REGION Network 16: Step7: Request Take Photos and Calculate Again When ROS Error | PLC Status Word:111 0r 112
   RUNG wire#powerrail
      Contact( #High )
      Contact( "DB2500 Visual Chiseling".VisualChiselingMode )
      Contact( "DB2500 Visual Chiseling".VisualCameraStart )
      wire#w1
      { S7_Templates := "SrcType := Int" } EQ_Contact(in1 := "DB2500 Visual Chiseling".RosErrorNum, in2 := 1)
      P_Trig( "DB2500 Visual Chiseling".Pulse[9] )
      Move(in := 111, out1 => "DB2100 Modbus Value"."PLC Para"."Status Word")
   END_RUNG
   RUNG wire#w1
      { S7_Templates := "SrcType := Int" } EQ_Contact(in1 := "DB2500 Visual Chiseling".RosErrorNum, in2 := 2)
      P_Trig( "DB2500 Visual Chiseling".Pulse[10] )
      Move(in := 112, out1 => "DB2100 Modbus Value"."PLC Para"."Status Word")
   END_RUNG
   // the same network as SCL:
   #_w1 := #High AND "DB2500 Visual Chiseling".VisualChiselingMode AND "DB2500 Visual Chiseling".VisualCameraStart;
   #_w2 := #_w1 AND ("DB2500 Visual Chiseling".RosErrorNum = 1);
   #_w3 := #_w2 AND NOT "DB2500 Visual Chiseling".Pulse[9];   // rising edge
   "DB2500 Visual Chiseling".Pulse[9] := #_w2;
   IF #_w3 THEN "DB2100 Modbus Value"."PLC Para"."Status Word" := 111; END_IF;
   #_w4 := #_w1 AND ("DB2500 Visual Chiseling".RosErrorNum = 2);
   #_w5 := #_w4 AND NOT "DB2500 Visual Chiseling".Pulse[10];   // rising edge
   "DB2500 Visual Chiseling".Pulse[10] := #_w4;
   IF #_w5 THEN "DB2100 Modbus Value"."PLC Para"."Status Word" := 112; END_IF;
END_REGION

REGION Network 17: Step7: Stop Communication and SShutDown ROS If Erro Num Bigger Than 3 | PLC Status Word:105
   // Status 105: Send Shut Down Signal to ROS
   RUNG wire#powerrail
      Contact( #High )
      Contact( "DB2500 Visual Chiseling".VisualChiselingMode )
      Contact( "DB2500 Visual Chiseling".VisualCameraStart )
      { S7_Templates := "SrcType := Int" } GE_Contact(in1 := "DB2500 Visual Chiseling".RosErrorNum, in2 := 3)
      P_Trig( "DB2500 Visual Chiseling".Pulse[11] )
      wire#w1
      Move(in := 105, out1 => "DB2100 Modbus Value"."PLC Para"."Status Word")
   END_RUNG
   RUNG wire#w1
      S_Coil( "DB2500 Visual Chiseling".ROSCalculationFault )
      R_Coil( "DB2500 Visual Chiseling".VisualCameraStart )
   END_RUNG
   // the same network as SCL:
   #_w1 := #High AND "DB2500 Visual Chiseling".VisualChiselingMode AND "DB2500 Visual Chiseling".VisualCameraStart AND ("DB2500 Visual Chiseling".RosErrorNum >= 3);
   #_w2 := #_w1 AND NOT "DB2500 Visual Chiseling".Pulse[11];   // rising edge
   "DB2500 Visual Chiseling".Pulse[11] := #_w1;
   IF #_w2 THEN
       "DB2100 Modbus Value"."PLC Para"."Status Word" := 105;
       "DB2500 Visual Chiseling".ROSCalculationFault := TRUE;
       "DB2500 Visual Chiseling".VisualCameraStart := FALSE;
   END_IF;
END_REGION

REGION Network 18: Step8: Auto Close Camera Protective Cover | PLC Status Word:130
   "Timer30_ChiselStepEnd".TON(IN := #High AND "DB2500 Visual Chiseling".VisualChiselingMode AND "DB2500 Visual Chiseling".VisualCameraStart AND (("DB2100 Modbus Value"."PLC Para"."Status Word" = 120) OR "DB2500 Visual Chiseling".ROSCalculationFault),
                           PT := T#0.2s);
   IF "Timer30_ChiselStepEnd".Q THEN "DB2100 Modbus Value"."PLC Para"."Status Word" := 130; END_IF;
END_REGION

REGION Network 19: Step9: Visual Chiseling Camera Function Completed
   // Robot: IN[80]   PLC :DB720.DBX2.0  VisualChiseling  Camera Function  Completion Signal
   RUNG wire#powerrail
      Contact( #High )
      Contact( "DB2500 Visual Chiseling".VisualChiselingMode )
      Contact( "DB2500 Visual Chiseling".VisualCameraStart )
      { S7_Templates := "SrcType := Word" } EQ_Contact(in1 := "DB2100 Modbus Value"."PLC Para"."Status Word", in2 := 130)
      P_Trig( "DB2500 Visual Chiseling".Pulse[12] )
      wire#w1
      Move(in := 0, out1 => "DB2500 Visual Chiseling".RosErrorNum)
   END_RUNG
   RUNG wire#w1
      R_Coil( "DB2500 Visual Chiseling".VisualCameraStart )
      S_Coil( "DB2500 Visual Chiseling".VisualCameraEnd )
      R_Coil( "QCamCoverExt" )
      S_Coil( "QCamCoverRet" )
   END_RUNG
   // the same network as SCL:
   #_w1 := #High AND "DB2500 Visual Chiseling".VisualChiselingMode AND "DB2500 Visual Chiseling".VisualCameraStart AND ("DB2100 Modbus Value"."PLC Para"."Status Word" = 130);
   #_w2 := #_w1 AND NOT "DB2500 Visual Chiseling".Pulse[12];   // rising edge
   "DB2500 Visual Chiseling".Pulse[12] := #_w1;
   IF #_w2 THEN
       "DB2500 Visual Chiseling".RosErrorNum := 0;
       "DB2500 Visual Chiseling".VisualCameraStart := FALSE;
       "DB2500 Visual Chiseling".VisualCameraEnd := TRUE;
       "QCamCoverExt" := FALSE;
       "QCamCoverRet" := TRUE;
   END_IF;
END_REGION

REGION Network 20: Step9.1 : Send Visual Chiseling Function Completion Signal to Robot.
   // Robot: IN[80]   PLC :DB720.DBX2.0  VisualChiseling  Camera Function  Completion Signal
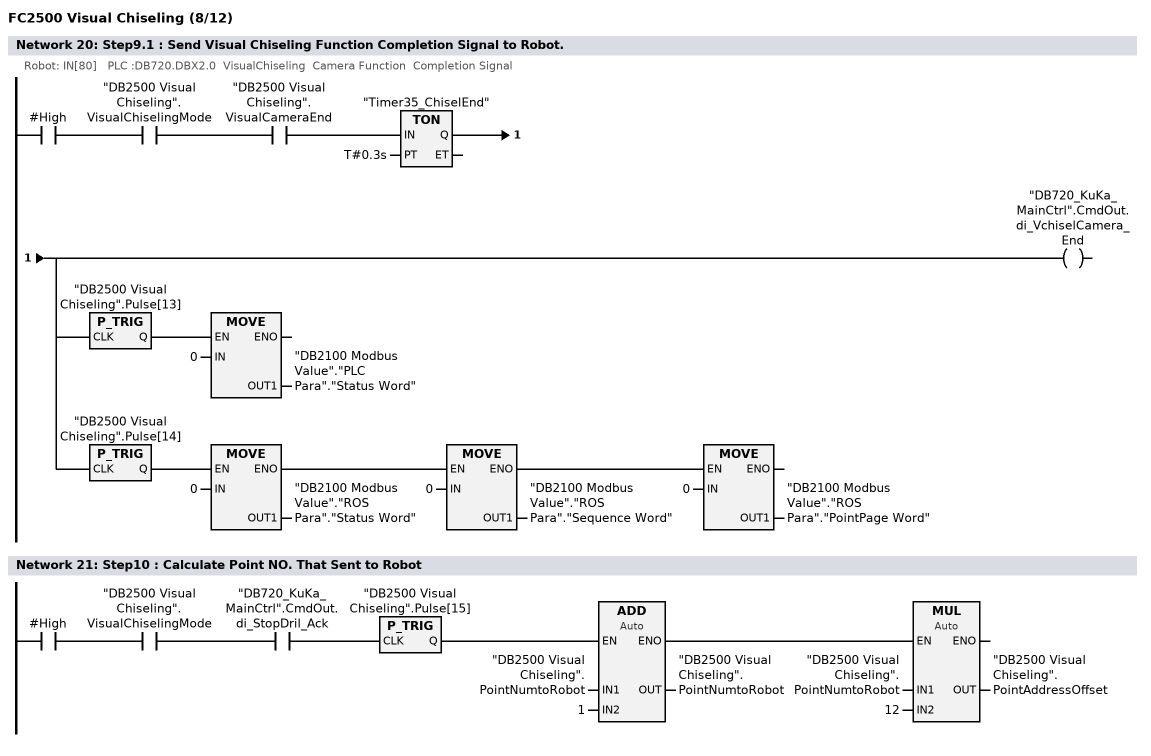
   "Timer35_ChiselEnd".TON(IN := #High AND "DB2500 Visual Chiseling".VisualChiselingMode AND "DB2500 Visual Chiseling".VisualCameraEnd,
                           PT := T#0.3s);
   "DB720_KuKa_MainCtrl".CmdOut.di_VchiselCamera_End := "Timer35_ChiselEnd".Q;
   #_w1 := "Timer35_ChiselEnd".Q AND NOT "DB2500 Visual Chiseling".Pulse[13];   // rising edge
   "DB2500 Visual Chiseling".Pulse[13] := "Timer35_ChiselEnd".Q;
   IF #_w1 THEN "DB2100 Modbus Value"."PLC Para"."Status Word" := 0; END_IF;
   #_w2 := "Timer35_ChiselEnd".Q AND NOT "DB2500 Visual Chiseling".Pulse[14];   // rising edge
   "DB2500 Visual Chiseling".Pulse[14] := "Timer35_ChiselEnd".Q;
   IF #_w2 THEN
       "DB2100 Modbus Value"."ROS Para"."Status Word" := 0;
       "DB2100 Modbus Value"."ROS Para"."Sequence Word" := 0;
       "DB2100 Modbus Value"."ROS Para"."PointPage Word" := 0;
   END_IF;
END_REGION

REGION Network 21: Step10 : Calculate Point NO. That Sent to Robot
   RUNG wire#powerrail
      Contact( #High )
      Contact( "DB2500 Visual Chiseling".VisualChiselingMode )
      Contact( "DB720_KuKa_MainCtrl".CmdOut.di_StopDril_Ack )
      P_Trig( "DB2500 Visual Chiseling".Pulse[15] )
      Add(in1 := "DB2500 Visual Chiseling".PointNumtoRobot, in2 := 1, out => "DB2500 Visual Chiseling".PointNumtoRobot)
      Mul(in1 := "DB2500 Visual Chiseling".PointNumtoRobot, in2 := 12, out => "DB2500 Visual Chiseling".PointAddressOffset)
   END_RUNG
   // the same network as SCL:
   #_w1 := #High AND "DB2500 Visual Chiseling".VisualChiselingMode AND "DB720_KuKa_MainCtrl".CmdOut.di_StopDril_Ack;
   #_w2 := #_w1 AND NOT "DB2500 Visual Chiseling".Pulse[15];   // rising edge
   "DB2500 Visual Chiseling".Pulse[15] := #_w1;
   IF #_w2 THEN
       "DB2500 Visual Chiseling".PointNumtoRobot := "DB2500 Visual Chiseling".PointNumtoRobot + 1;
       "DB2500 Visual Chiseling".PointAddressOffset := "DB2500 Visual Chiseling".PointNumtoRobot * 12;
   END_IF;
END_REGION

REGION Network 22 (SCL): Step11: Move Current Chiseling Point to Offset Value. (SCL)
   // byteOffset_dest Should Be Changed wehn
   IF "DB2500 Visual Chiseling".VisualCameraEnd = TRUE THEN
       POKE_BLK(area_src := 16#84,
                dbNumber_src := 2300,
                byteOffset_src := "DB2500 Visual Chiseling".PointAddressOffset,
                area_dest := 16#84,
                dbNumber_dest := 2500,
                byteOffset_dest := 38,
                count := 12);
   END_IF;
END_REGION

REGION Network 23: Step12: Offset Value Format From Word To Real
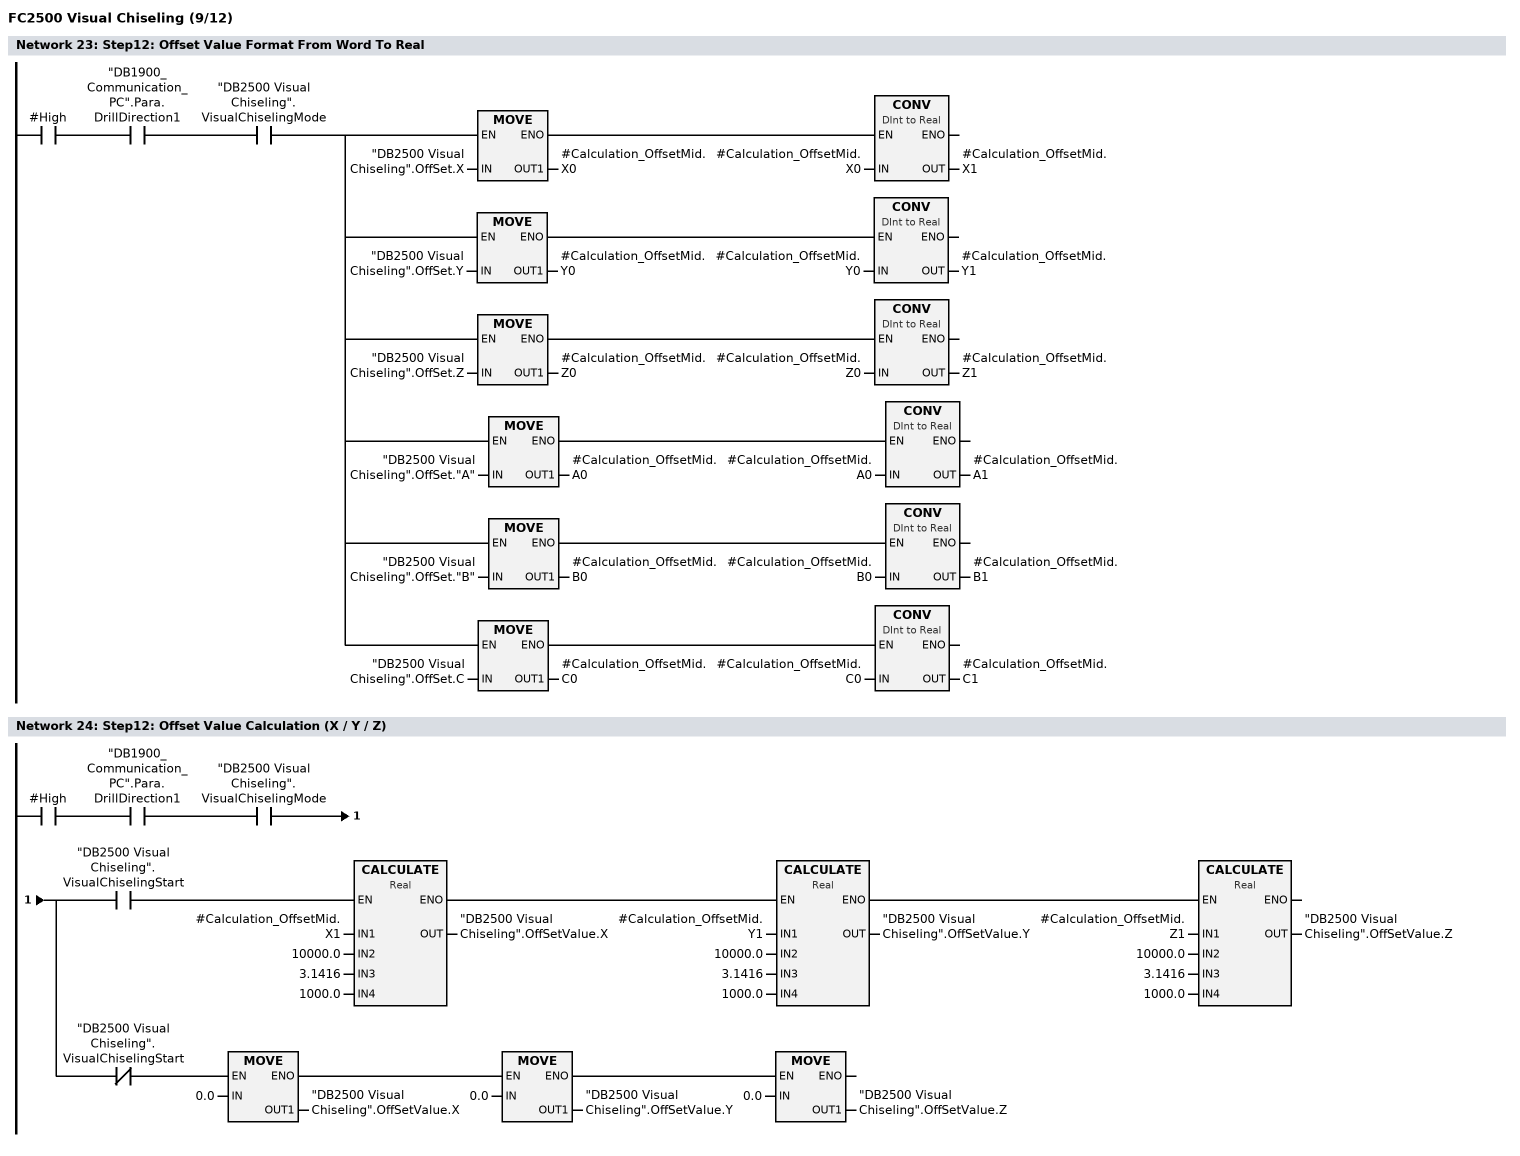
   RUNG wire#powerrail
      Contact( #High )
      Contact( "DB1900_Communication_PC".Para.DrillDirection1 )
      Contact( "DB2500 Visual Chiseling".VisualChiselingMode )
      wire#w1
      Move(in := "DB2500 Visual Chiseling".OffSet.X, out1 => #Calculation_OffsetMid.X0)
      { S7_Templates := "[SrcType := DInt, DestType := Real]" } Convert(in := #Calculation_OffsetMid.X0, out => #Calculation_OffsetMid.X1)
   END_RUNG
   RUNG wire#w1
      Move(in := "DB2500 Visual Chiseling".OffSet.Y, out1 => #Calculation_OffsetMid.Y0)
      { S7_Templates := "[SrcType := DInt, DestType := Real]" } Convert(in := #Calculation_OffsetMid.Y0, out => #Calculation_OffsetMid.Y1)
   END_RUNG
   RUNG wire#w1
      Move(in := "DB2500 Visual Chiseling".OffSet.Z, out1 => #Calculation_OffsetMid.Z0)
      { S7_Templates := "[SrcType := DInt, DestType := Real]" } Convert(in := #Calculation_OffsetMid.Z0, out => #Calculation_OffsetMid.Z1)
   END_RUNG
   RUNG wire#w1
      Move(in := "DB2500 Visual Chiseling".OffSet."A", out1 => #Calculation_OffsetMid.A0)
      { S7_Templates := "[SrcType := DInt, DestType := Real]" } Convert(in := #Calculation_OffsetMid.A0, out => #Calculation_OffsetMid.A1)
   END_RUNG
   RUNG wire#w1
      Move(in := "DB2500 Visual Chiseling".OffSet."B", out1 => #Calculation_OffsetMid.B0)
      { S7_Templates := "[SrcType := DInt, DestType := Real]" } Convert(in := #Calculation_OffsetMid.B0, out => #Calculation_OffsetMid.B1)
   END_RUNG
   RUNG wire#w1
      Move(in := "DB2500 Visual Chiseling".OffSet.C, out1 => #Calculation_OffsetMid.C0)
      { S7_Templates := "[SrcType := DInt, DestType := Real]" } Convert(in := #Calculation_OffsetMid.C0, out => #Calculation_OffsetMid.C1)
   END_RUNG
   // the same network as SCL:
   IF #High AND "DB1900_Communication_PC".Para.DrillDirection1 AND "DB2500 Visual Chiseling".VisualChiselingMode THEN
       #Calculation_OffsetMid.X0 := "DB2500 Visual Chiseling".OffSet.X;
       #Calculation_OffsetMid.X1 := DINT_TO_REAL(#Calculation_OffsetMid.X0);
       #Calculation_OffsetMid.Y0 := "DB2500 Visual Chiseling".OffSet.Y;
       #Calculation_OffsetMid.Y1 := DINT_TO_REAL(#Calculation_OffsetMid.Y0);
       #Calculation_OffsetMid.Z0 := "DB2500 Visual Chiseling".OffSet.Z;
       #Calculation_OffsetMid.Z1 := DINT_TO_REAL(#Calculation_OffsetMid.Z0);
       #Calculation_OffsetMid.A0 := "DB2500 Visual Chiseling".OffSet."A";
       #Calculation_OffsetMid.A1 := DINT_TO_REAL(#Calculation_OffsetMid.A0);
       #Calculation_OffsetMid.B0 := "DB2500 Visual Chiseling".OffSet."B";
       #Calculation_OffsetMid.B1 := DINT_TO_REAL(#Calculation_OffsetMid.B0);
       #Calculation_OffsetMid.C0 := "DB2500 Visual Chiseling".OffSet.C;
       #Calculation_OffsetMid.C1 := DINT_TO_REAL(#Calculation_OffsetMid.C0);
   END_IF;
END_REGION

REGION Network 24: Step12: Offset Value Calculation (X / Y / Z)
   RUNG wire#powerrail
      Contact( #High )
      Contact( "DB1900_Communication_PC".Para.DrillDirection1 )
      Contact( "DB2500 Visual Chiseling".VisualChiselingMode )
      wire#w1
      Contact( "DB2500 Visual Chiseling".VisualChiselingStart )
      { S7_Templates := "SrcType := Real"; S7_Expression := "( IN1 / IN2 - IN3 ) * IN4" } Calculate(in1 := #Calculation_OffsetMid.X1, in2 := 10000.0, in3 := 3.1416, in4 := 1000.0, out => "DB2500 Visual Chiseling".OffSetValue.X)
      { S7_Templates := "SrcType := Real"; S7_Expression := "( IN1 / IN2 - IN3 ) * IN4" } Calculate(in1 := #Calculation_OffsetMid.Y1, in2 := 10000.0, in3 := 3.1416, in4 := 1000.0, out => "DB2500 Visual Chiseling".OffSetValue.Y)
      { S7_Templates := "SrcType := Real"; S7_Expression := "( IN1 / IN2 - IN3 ) * IN4" } Calculate(in1 := #Calculation_OffsetMid.Z1, in2 := 10000.0, in3 := 3.1416, in4 := 1000.0, out => "DB2500 Visual Chiseling".OffSetValue.Z)
   END_RUNG
   RUNG wire#w1
      I_Contact( "DB2500 Visual Chiseling".VisualChiselingStart )
      Move(in := 0.0, out1 => "DB2500 Visual Chiseling".OffSetValue.X)
      Move(in := 0.0, out1 => "DB2500 Visual Chiseling".OffSetValue.Y)
      Move(in := 0.0, out1 => "DB2500 Visual Chiseling".OffSetValue.Z)
   END_RUNG
   // the same network as SCL:
   #_w1 := #High AND "DB1900_Communication_PC".Para.DrillDirection1 AND "DB2500 Visual Chiseling".VisualChiselingMode;
   IF #_w1 AND "DB2500 Visual Chiseling".VisualChiselingStart THEN
       "DB2500 Visual Chiseling".OffSetValue.X := ( #Calculation_OffsetMid.X1 / 10000.0 - 3.1416 ) * 1000.0;
       "DB2500 Visual Chiseling".OffSetValue.Y := ( #Calculation_OffsetMid.Y1 / 10000.0 - 3.1416 ) * 1000.0;
       "DB2500 Visual Chiseling".OffSetValue.Z := ( #Calculation_OffsetMid.Z1 / 10000.0 - 3.1416 ) * 1000.0;
   END_IF;
   IF #_w1 AND NOT "DB2500 Visual Chiseling".VisualChiselingStart THEN
       "DB2500 Visual Chiseling".OffSetValue.X := 0.0;
       "DB2500 Visual Chiseling".OffSetValue.Y := 0.0;
       "DB2500 Visual Chiseling".OffSetValue.Z := 0.0;
   END_IF;
END_REGION

REGION Network 25: Step13: Offset Value Calculation (A / B / C)
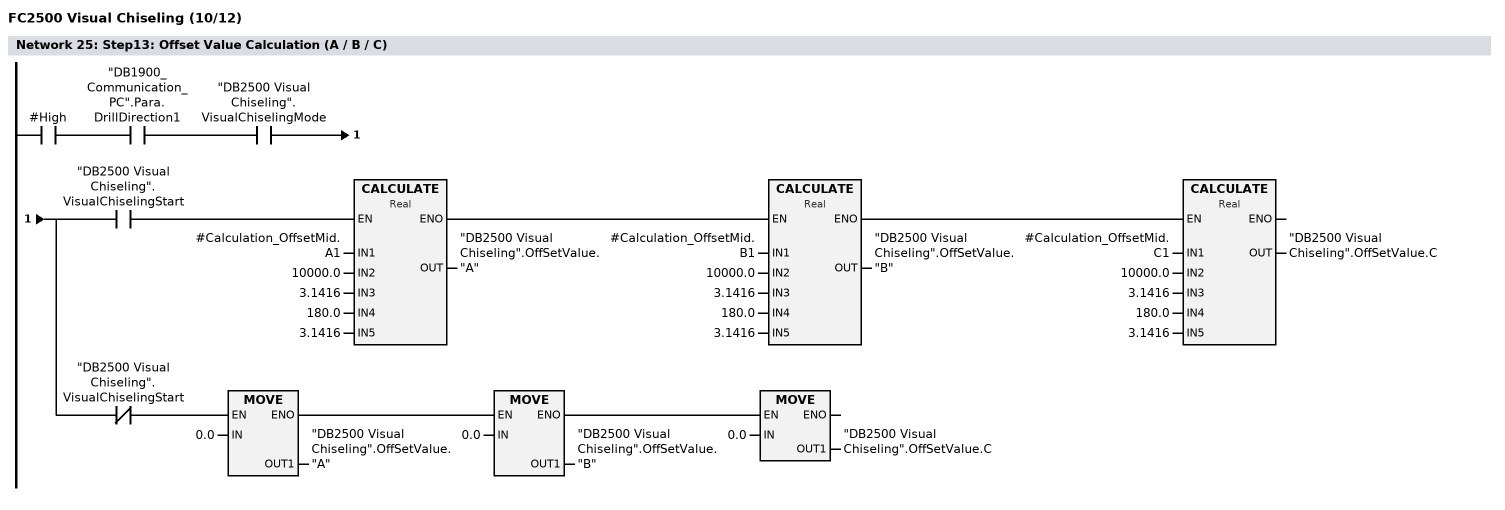
   RUNG wire#powerrail
      Contact( #High )
      Contact( "DB1900_Communication_PC".Para.DrillDirection1 )
      Contact( "DB2500 Visual Chiseling".VisualChiselingMode )
      wire#w1
      Contact( "DB2500 Visual Chiseling".VisualChiselingStart )
      { S7_Templates := "SrcType := Real"; S7_Expression := "( ( IN1 / IN2 - IN3 ) * IN4 ) / IN5" } Calculate(in1 := #Calculation_OffsetMid.A1, in2 := 10000.0, in3 := 3.1416, in4 := 180.0, in5 := 3.1416, out => "DB2500 Visual Chiseling".OffSetValue."A")
      { S7_Templates := "SrcType := Real"; S7_Expression := "( ( IN1 / IN2 - IN3 ) * IN4 ) / IN5" } Calculate(in1 := #Calculation_OffsetMid.B1, in2 := 10000.0, in3 := 3.1416, in4 := 180.0, in5 := 3.1416, out => "DB2500 Visual Chiseling".OffSetValue."B")
      { S7_Templates := "SrcType := Real"; S7_Expression := "( ( IN1 / IN2 - IN3 ) * IN4 ) / IN5" } Calculate(in1 := #Calculation_OffsetMid.C1, in2 := 10000.0, in3 := 3.1416, in4 := 180.0, in5 := 3.1416, out => "DB2500 Visual Chiseling".OffSetValue.C)
   END_RUNG
   RUNG wire#w1
      I_Contact( "DB2500 Visual Chiseling".VisualChiselingStart )
      Move(in := 0.0, out1 => "DB2500 Visual Chiseling".OffSetValue."A")
      Move(in := 0.0, out1 => "DB2500 Visual Chiseling".OffSetValue."B")
      Move(in := 0.0, out1 => "DB2500 Visual Chiseling".OffSetValue.C)
   END_RUNG
   // the same network as SCL:
   #_w1 := #High AND "DB1900_Communication_PC".Para.DrillDirection1 AND "DB2500 Visual Chiseling".VisualChiselingMode;
   IF #_w1 AND "DB2500 Visual Chiseling".VisualChiselingStart THEN
       "DB2500 Visual Chiseling".OffSetValue."A" := ( ( #Calculation_OffsetMid.A1 / 10000.0 - 3.1416 ) * 180.0 ) / 3.1416;
       "DB2500 Visual Chiseling".OffSetValue."B" := ( ( #Calculation_OffsetMid.B1 / 10000.0 - 3.1416 ) * 180.0 ) / 3.1416;
       "DB2500 Visual Chiseling".OffSetValue.C := ( ( #Calculation_OffsetMid.C1 / 10000.0 - 3.1416 ) * 180.0 ) / 3.1416;
   END_IF;
   IF #_w1 AND NOT "DB2500 Visual Chiseling".VisualChiselingStart THEN
       "DB2500 Visual Chiseling".OffSetValue."A" := 0.0;
       "DB2500 Visual Chiseling".OffSetValue."B" := 0.0;
       "DB2500 Visual Chiseling".OffSetValue.C := 0.0;
   END_IF;
END_REGION

REGION Network 26: Step14: Transfer Offset Value to Robot
   // Added by WXY 20220618.  DBD720.DBD36: gi_OffSetA;  DBD720.DBD40: gi_OffSetB;   DBD720.DBD44: gi_OffSetC
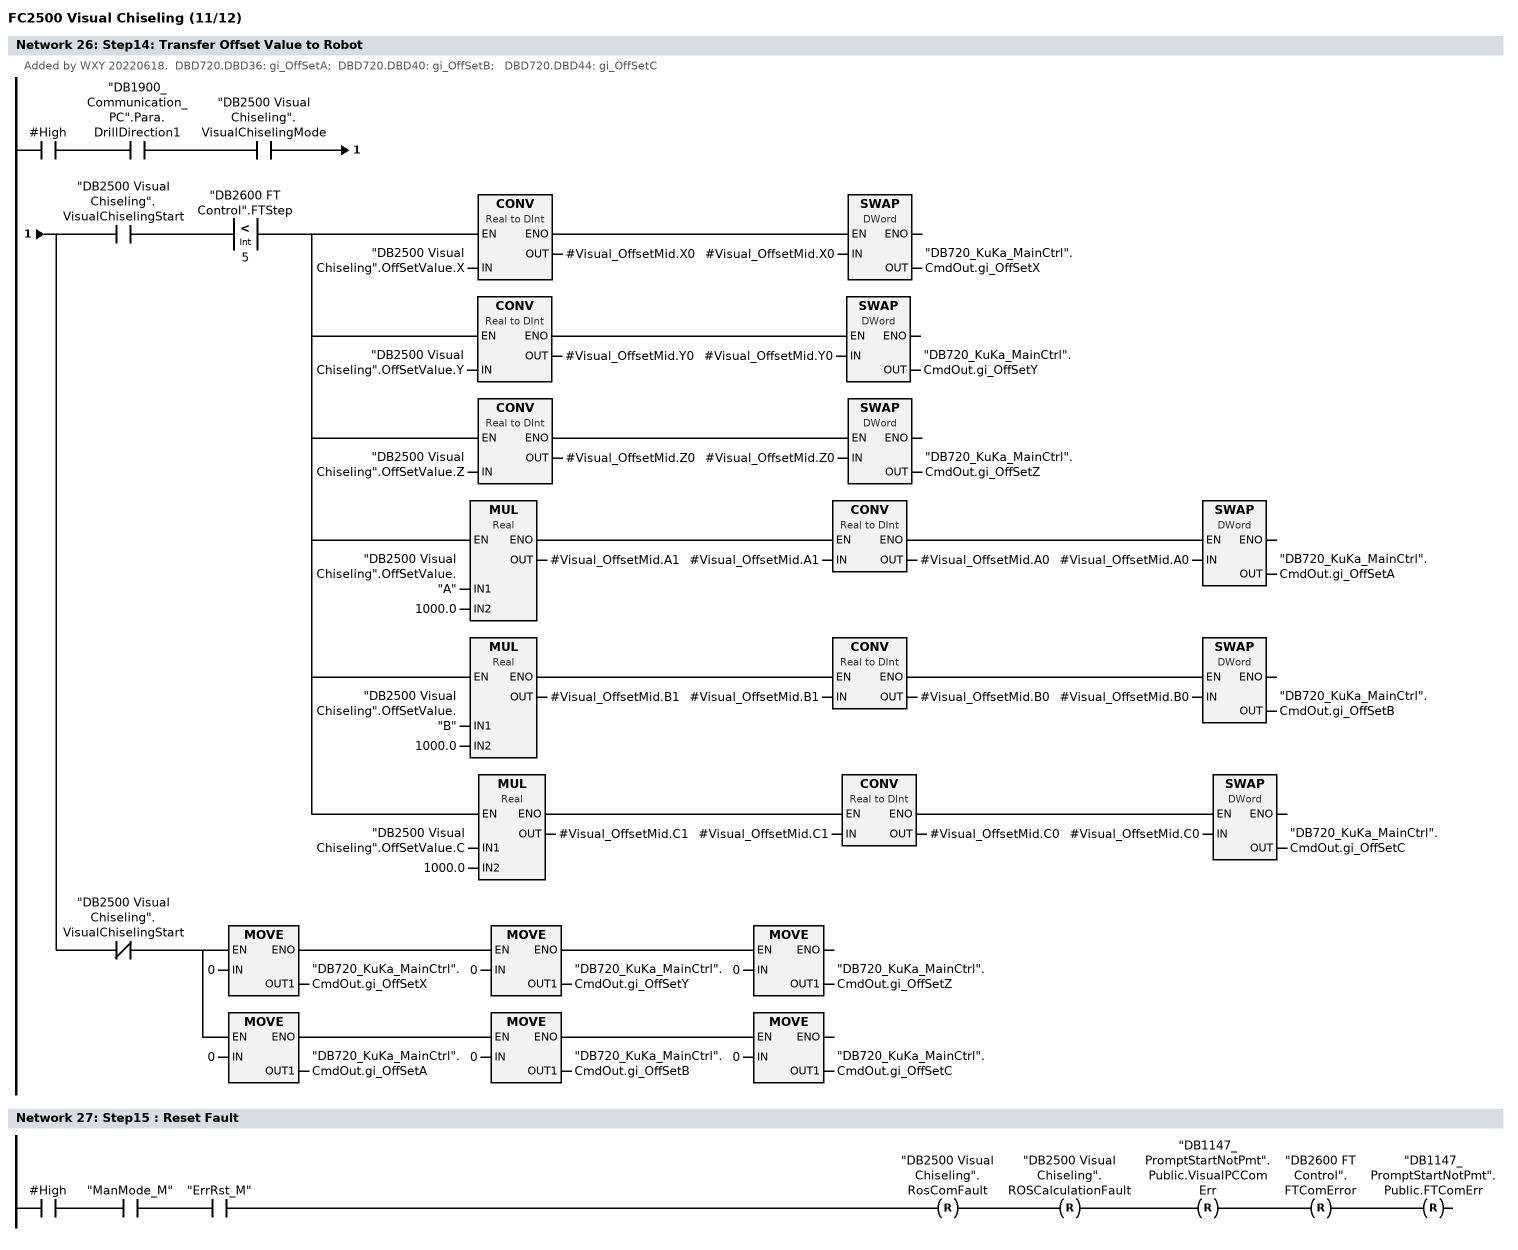
   #_w1 := #High AND "DB1900_Communication_PC".Para.DrillDirection1 AND "DB2500 Visual Chiseling".VisualChiselingMode;
   IF #_w1 AND "DB2500 Visual Chiseling".VisualChiselingStart AND ("DB2600 FT Control".FTStep < 5) THEN
       #Visual_OffsetMid.X0 := REAL_TO_DINT("DB2500 Visual Chiseling".OffSetValue.X);
       "DB720_KuKa_MainCtrl".CmdOut.gi_OffSetX := SWAP(#Visual_OffsetMid.X0);
       #Visual_OffsetMid.Y0 := REAL_TO_DINT("DB2500 Visual Chiseling".OffSetValue.Y);
       "DB720_KuKa_MainCtrl".CmdOut.gi_OffSetY := SWAP(#Visual_OffsetMid.Y0);
       #Visual_OffsetMid.Z0 := REAL_TO_DINT("DB2500 Visual Chiseling".OffSetValue.Z);
       "DB720_KuKa_MainCtrl".CmdOut.gi_OffSetZ := SWAP(#Visual_OffsetMid.Z0);
       #Visual_OffsetMid.A1 := "DB2500 Visual Chiseling".OffSetValue."A" * 1000.0;
       #Visual_OffsetMid.A0 := REAL_TO_DINT(#Visual_OffsetMid.A1);
       "DB720_KuKa_MainCtrl".CmdOut.gi_OffSetA := SWAP(#Visual_OffsetMid.A0);
       #Visual_OffsetMid.B1 := "DB2500 Visual Chiseling".OffSetValue."B" * 1000.0;
       #Visual_OffsetMid.B0 := REAL_TO_DINT(#Visual_OffsetMid.B1);
       "DB720_KuKa_MainCtrl".CmdOut.gi_OffSetB := SWAP(#Visual_OffsetMid.B0);
       #Visual_OffsetMid.C1 := "DB2500 Visual Chiseling".OffSetValue.C * 1000.0;
       #Visual_OffsetMid.C0 := REAL_TO_DINT(#Visual_OffsetMid.C1);
       "DB720_KuKa_MainCtrl".CmdOut.gi_OffSetC := SWAP(#Visual_OffsetMid.C0);
   END_IF;
   IF #_w1 AND NOT "DB2500 Visual Chiseling".VisualChiselingStart THEN
       "DB720_KuKa_MainCtrl".CmdOut.gi_OffSetX := 0;
       "DB720_KuKa_MainCtrl".CmdOut.gi_OffSetY := 0;
       "DB720_KuKa_MainCtrl".CmdOut.gi_OffSetZ := 0;
       "DB720_KuKa_MainCtrl".CmdOut.gi_OffSetA := 0;
       "DB720_KuKa_MainCtrl".CmdOut.gi_OffSetB := 0;
       "DB720_KuKa_MainCtrl".CmdOut.gi_OffSetC := 0;
   END_IF;
END_REGION

REGION Network 27: Step15 : Reset Fault
   RUNG wire#powerrail
      Contact( #High )
      Contact( "ManMode_M" )
      Contact( "ErrRst_M" )
      R_Coil( "DB2500 Visual Chiseling".RosComFault )
      R_Coil( "DB2500 Visual Chiseling".ROSCalculationFault )
      R_Coil( "DB1147_PromptStartNotPmt".Public.VisualPCComErr )
      R_Coil( "DB2600 FT Control".FTComError )
      R_Coil( "DB1147_PromptStartNotPmt".Public.FTComErr )
   END_RUNG
   // the same network as SCL:
   IF #High AND "ManMode_M" AND "ErrRst_M" THEN
       "DB2500 Visual Chiseling".RosComFault := FALSE;
       "DB2500 Visual Chiseling".ROSCalculationFault := FALSE;
       "DB1147_PromptStartNotPmt".Public.VisualPCComErr := FALSE;
       "DB2600 FT Control".FTComError := FALSE;
       "DB1147_PromptStartNotPmt".Public.FTComErr := FALSE;
   END_IF;
END_REGION

REGION Network 28: ################# Cal Cam Round #################
END_REGION

REGION Network 29: Reset Camera Round
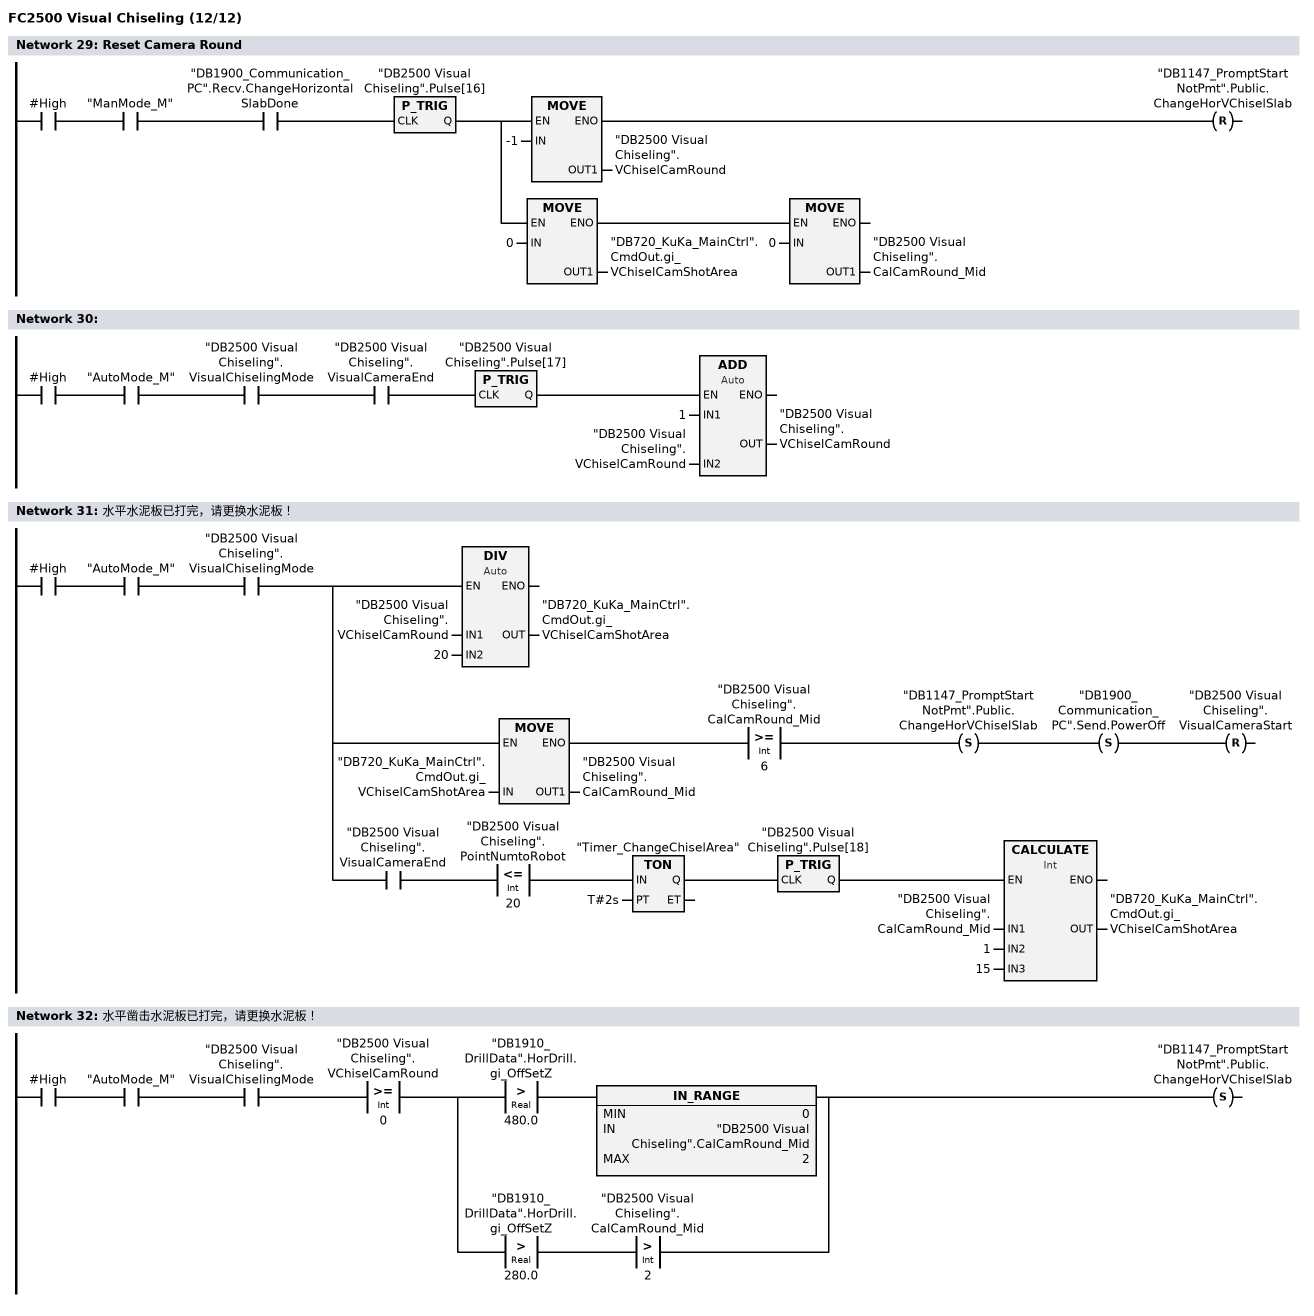
   RUNG wire#powerrail
      Contact( #High )
      Contact( "ManMode_M" )
      Contact( "DB1900_Communication_PC".Recv.ChangeHorizontalSlabDone )
      P_Trig( "DB2500 Visual Chiseling".Pulse[16] )
      wire#w1
      Move(in := -1, out1 => "DB2500 Visual Chiseling".VChiselCamRound)
      R_Coil( "DB1147_PromptStartNotPmt".Public.ChangeHorVChiselSlab )
   END_RUNG
   RUNG wire#w1
      Move(in := 0, out1 => "DB720_KuKa_MainCtrl".CmdOut.gi_VChiselCamShotArea)
      Move(in := 0, out1 => "DB2500 Visual Chiseling".CalCamRound_Mid)
   END_RUNG
   // the same network as SCL:
   #_w1 := #High AND "ManMode_M" AND "DB1900_Communication_PC".Recv.ChangeHorizontalSlabDone;
   #_w2 := #_w1 AND NOT "DB2500 Visual Chiseling".Pulse[16];   // rising edge
   "DB2500 Visual Chiseling".Pulse[16] := #_w1;
   IF #_w2 THEN
       "DB2500 Visual Chiseling".VChiselCamRound := -1;
       "DB1147_PromptStartNotPmt".Public.ChangeHorVChiselSlab := FALSE;
       "DB720_KuKa_MainCtrl".CmdOut.gi_VChiselCamShotArea := 0;
       "DB2500 Visual Chiseling".CalCamRound_Mid := 0;
   END_IF;
END_REGION

REGION Network 30
   RUNG wire#powerrail
      Contact( #High )
      Contact( "AutoMode_M" )
      Contact( "DB2500 Visual Chiseling".VisualChiselingMode )
      Contact( "DB2500 Visual Chiseling".VisualCameraEnd )
      P_Trig( "DB2500 Visual Chiseling".Pulse[17] )
      Add(in1 := 1, in2 := "DB2500 Visual Chiseling".VChiselCamRound, out => "DB2500 Visual Chiseling".VChiselCamRound)
   END_RUNG
   // the same network as SCL:
   #_w1 := #High AND "AutoMode_M" AND "DB2500 Visual Chiseling".VisualChiselingMode AND "DB2500 Visual Chiseling".VisualCameraEnd;
   #_w2 := #_w1 AND NOT "DB2500 Visual Chiseling".Pulse[17];   // rising edge
   "DB2500 Visual Chiseling".Pulse[17] := #_w1;
   IF #_w2 THEN
       "DB2500 Visual Chiseling".VChiselCamRound := 1 + "DB2500 Visual Chiseling".VChiselCamRound;
   END_IF;
END_REGION

REGION Network 31: 水平水泥板已打完，请更换水泥板！
   #_w1 := #High AND "AutoMode_M" AND "DB2500 Visual Chiseling".VisualChiselingMode;
   IF #_w1 THEN
       "DB720_KuKa_MainCtrl".CmdOut.gi_VChiselCamShotArea := "DB2500 Visual Chiseling".VChiselCamRound / 20;
       "DB2500 Visual Chiseling".CalCamRound_Mid := "DB720_KuKa_MainCtrl".CmdOut.gi_VChiselCamShotArea;
   END_IF;
   IF #_w1 AND ("DB2500 Visual Chiseling".CalCamRound_Mid >= 6) THEN
       "DB1147_PromptStartNotPmt".Public.ChangeHorVChiselSlab := TRUE;
       "DB1900_Communication_PC".Send.PowerOff := TRUE;
       "DB2500 Visual Chiseling".VisualCameraStart := FALSE;
   END_IF;
   "Timer_ChangeChiselArea".TON(IN := #_w1 AND "DB2500 Visual Chiseling".VisualCameraEnd AND ("DB2500 Visual Chiseling".PointNumtoRobot <= 20),
                           PT := T#2s);
   #_w2 := "Timer_ChangeChiselArea".Q AND NOT "DB2500 Visual Chiseling".Pulse[18];   // rising edge
   "DB2500 Visual Chiseling".Pulse[18] := "Timer_ChangeChiselArea".Q;
   IF #_w2 THEN
       "DB720_KuKa_MainCtrl".CmdOut.gi_VChiselCamShotArea := ("DB2500 Visual Chiseling".CalCamRound_Mid+1)*15;
   END_IF;
END_REGION

REGION Network 32: 水平凿击水泥板已打完，请更换水泥板！
   RUNG wire#powerrail
      Contact( #High )
      Contact( "AutoMode_M" )
      Contact( "DB2500 Visual Chiseling".VisualChiselingMode )
      { S7_Templates := "SrcType := Int" } GE_Contact(in1 := "DB2500 Visual Chiseling".VChiselCamRound, in2 := 0)
      wire#w1
      { S7_Templates := "SrcType := Real" } GT_Contact(in1 := "DB1910_DrillData".HorDrill.gi_OffSetZ, in2 := 480.0)
      { S7_Templates := "SrcType := Int" } InRange(min := 0, in := "DB2500 Visual Chiseling".CalCamRound_Mid, max := 2)
      wire#w2
      S_Coil( "DB1147_PromptStartNotPmt".Public.ChangeHorVChiselSlab )
   END_RUNG
   RUNG wire#w1
      { S7_Templates := "SrcType := Real" } GT_Contact(in1 := "DB1910_DrillData".HorDrill.gi_OffSetZ, in2 := 280.0)
      { S7_Templates := "SrcType := Int" } GT_Contact(in1 := "DB2500 Visual Chiseling".CalCamRound_Mid, in2 := 2)
   END_RUNG wire#w2
   // the same network as SCL:
   IF #High AND "AutoMode_M" AND "DB2500 Visual Chiseling".VisualChiselingMode AND ("DB2500 Visual Chiseling".VChiselCamRound >= 0) AND ((("DB1910_DrillData".HorDrill.gi_OffSetZ > 480.0) AND (0 <= "DB2500 Visual Chiseling".CalCamRound_Mid) AND ("DB2500 Visual Chiseling".CalCamRound_Mid <= 2)) OR (("DB1910_DrillData".HorDrill.gi_OffSetZ > 280.0) AND ("DB2500 Visual Chiseling".CalCamRound_Mid > 2))) THEN
       "DB1147_PromptStartNotPmt".Public.ChangeHorVChiselSlab := TRUE;
   END_IF;
END_REGION
END_FUNCTION

FUNCTION "FC2600 FT Control" : Void   // FC2600, LAD
{ S7_Optimized_Access := 'TRUE' }
VERSION : 0.1
   VAR_TEMP
      FT_Calib_Done : Bool;
      FT_Recv_Done : Bool;
      MV_Ret_Val : Int;
      TarPoint_REAL : Struct
         X : Real;
         Y : Real;
         Z : Real;
         "A" : Real;
         "B" : Real;
         C : Real;
      END_STRUCT;
      TarPoint_DINT : Struct
         X : DInt;
         Y : DInt;
         Z : DInt;
         "A" : DInt;
         "B" : DInt;
         C : DInt;
      END_STRUCT;
      TTT : Bool;
   END_VAR
   VAR_TEMP   // added for the SCL form of the ladder/FBD networks
      _w1 : Bool;
      _w2 : Bool;
      _w3 : Bool;
      _w4 : Bool;
      _w5 : Bool;
      _w6 : Bool;
      _w7 : Bool;
      _w8 : Bool;
   END_VAR
BEGIN

REGION Network 1: Step0: only activate in vchisel mode
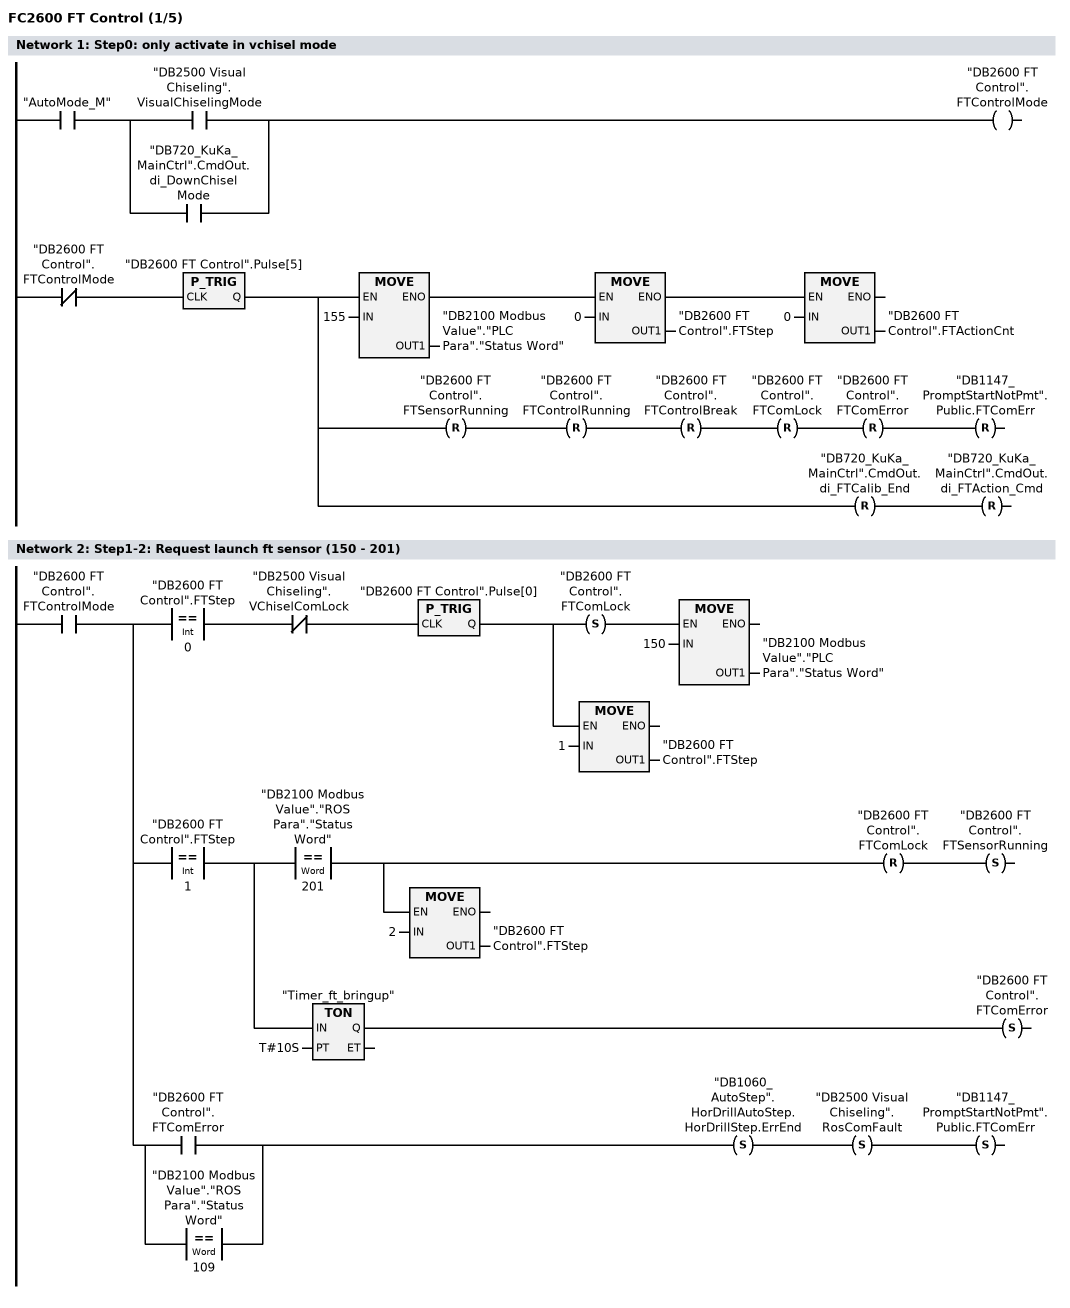
   RUNG wire#powerrail
      Contact( "AutoMode_M" )
      wire#w1
      Contact( "DB2500 Visual Chiseling".VisualChiselingMode )
      wire#w2
      Coil( "DB2600 FT Control".FTControlMode )
   END_RUNG
   RUNG wire#w1
      Contact( "DB720_KuKa_MainCtrl".CmdOut.di_DownChiselMode )
   END_RUNG wire#w2
   RUNG wire#powerrail
      I_Contact( "DB2600 FT Control".FTControlMode )
      P_Trig( "DB2600 FT Control".Pulse[5] )
      wire#w3
      Move(in := 155, out1 => "DB2100 Modbus Value"."PLC Para"."Status Word")
      Move(in := 0, out1 => "DB2600 FT Control".FTStep)
      Move(in := 0, out1 => "DB2600 FT Control".FTActionCnt)
   END_RUNG
   RUNG wire#w3
      R_Coil( "DB2600 FT Control".FTSensorRunning )
      R_Coil( "DB2600 FT Control".FTControlRunning )
      R_Coil( "DB2600 FT Control".FTControlBreak )
      R_Coil( "DB2600 FT Control".FTComLock )
      R_Coil( "DB2600 FT Control".FTComError )
      R_Coil( "DB1147_PromptStartNotPmt".Public.FTComErr )
   END_RUNG
   RUNG wire#w3
      R_Coil( "DB720_KuKa_MainCtrl".CmdOut.di_FTCalib_End )
      R_Coil( "DB720_KuKa_MainCtrl".CmdOut.di_FTAction_Cmd )
   END_RUNG
   // the same network as SCL:
   "DB2600 FT Control".FTControlMode := "AutoMode_M" AND ("DB2500 Visual Chiseling".VisualChiselingMode OR "DB720_KuKa_MainCtrl".CmdOut.di_DownChiselMode);
   #_w1 := NOT "DB2600 FT Control".FTControlMode AND NOT "DB2600 FT Control".Pulse[5];   // rising edge
   "DB2600 FT Control".Pulse[5] := NOT "DB2600 FT Control".FTControlMode;
   IF #_w1 THEN
       "DB2100 Modbus Value"."PLC Para"."Status Word" := 155;
       "DB2600 FT Control".FTStep := 0;
       "DB2600 FT Control".FTActionCnt := 0;
       "DB2600 FT Control".FTSensorRunning := FALSE;
       "DB2600 FT Control".FTControlRunning := FALSE;
       "DB2600 FT Control".FTControlBreak := FALSE;
       "DB2600 FT Control".FTComLock := FALSE;
       "DB2600 FT Control".FTComError := FALSE;
       "DB1147_PromptStartNotPmt".Public.FTComErr := FALSE;
       "DB720_KuKa_MainCtrl".CmdOut.di_FTCalib_End := FALSE;
       "DB720_KuKa_MainCtrl".CmdOut.di_FTAction_Cmd := FALSE;
   END_IF;
END_REGION

REGION Network 2: Step1-2: Request launch ft sensor (150 - 201)
   #_w1 := "DB2600 FT Control".FTControlMode AND ("DB2600 FT Control".FTStep = 0) AND NOT "DB2500 Visual Chiseling".VChiselComLock;
   #_w2 := #_w1 AND NOT "DB2600 FT Control".Pulse[0];   // rising edge
   "DB2600 FT Control".Pulse[0] := #_w1;
   IF #_w2 THEN
       "DB2600 FT Control".FTComLock := TRUE;
       "DB2100 Modbus Value"."PLC Para"."Status Word" := 150;
       "DB2600 FT Control".FTStep := 1;
   END_IF;
   #_w3 := "DB2600 FT Control".FTControlMode AND ("DB2600 FT Control".FTStep = 1);
   IF #_w3 AND ("DB2100 Modbus Value"."ROS Para"."Status Word" = 201) THEN
       "DB2600 FT Control".FTComLock := FALSE;
       "DB2600 FT Control".FTSensorRunning := TRUE;
       "DB2600 FT Control".FTStep := 2;
   END_IF;
   "Timer_ft_bringup".TON(IN := #_w3, PT := T#10S);
   IF "Timer_ft_bringup".Q THEN "DB2600 FT Control".FTComError := TRUE; END_IF;
   IF "DB2600 FT Control".FTControlMode AND ("DB2600 FT Control".FTComError OR ("DB2100 Modbus Value"."ROS Para"."Status Word" = 109)) THEN
       "DB1060_AutoStep".HorDrillAutoStep.HorDrillStep.ErrEnd := TRUE;
       "DB2500 Visual Chiseling".RosComFault := TRUE;
       "DB1147_PromptStartNotPmt".Public.FTComErr := TRUE;
   END_IF;
END_REGION

REGION Network 3: Step3-4: Ruquest calib ft sensor (160 - 202)
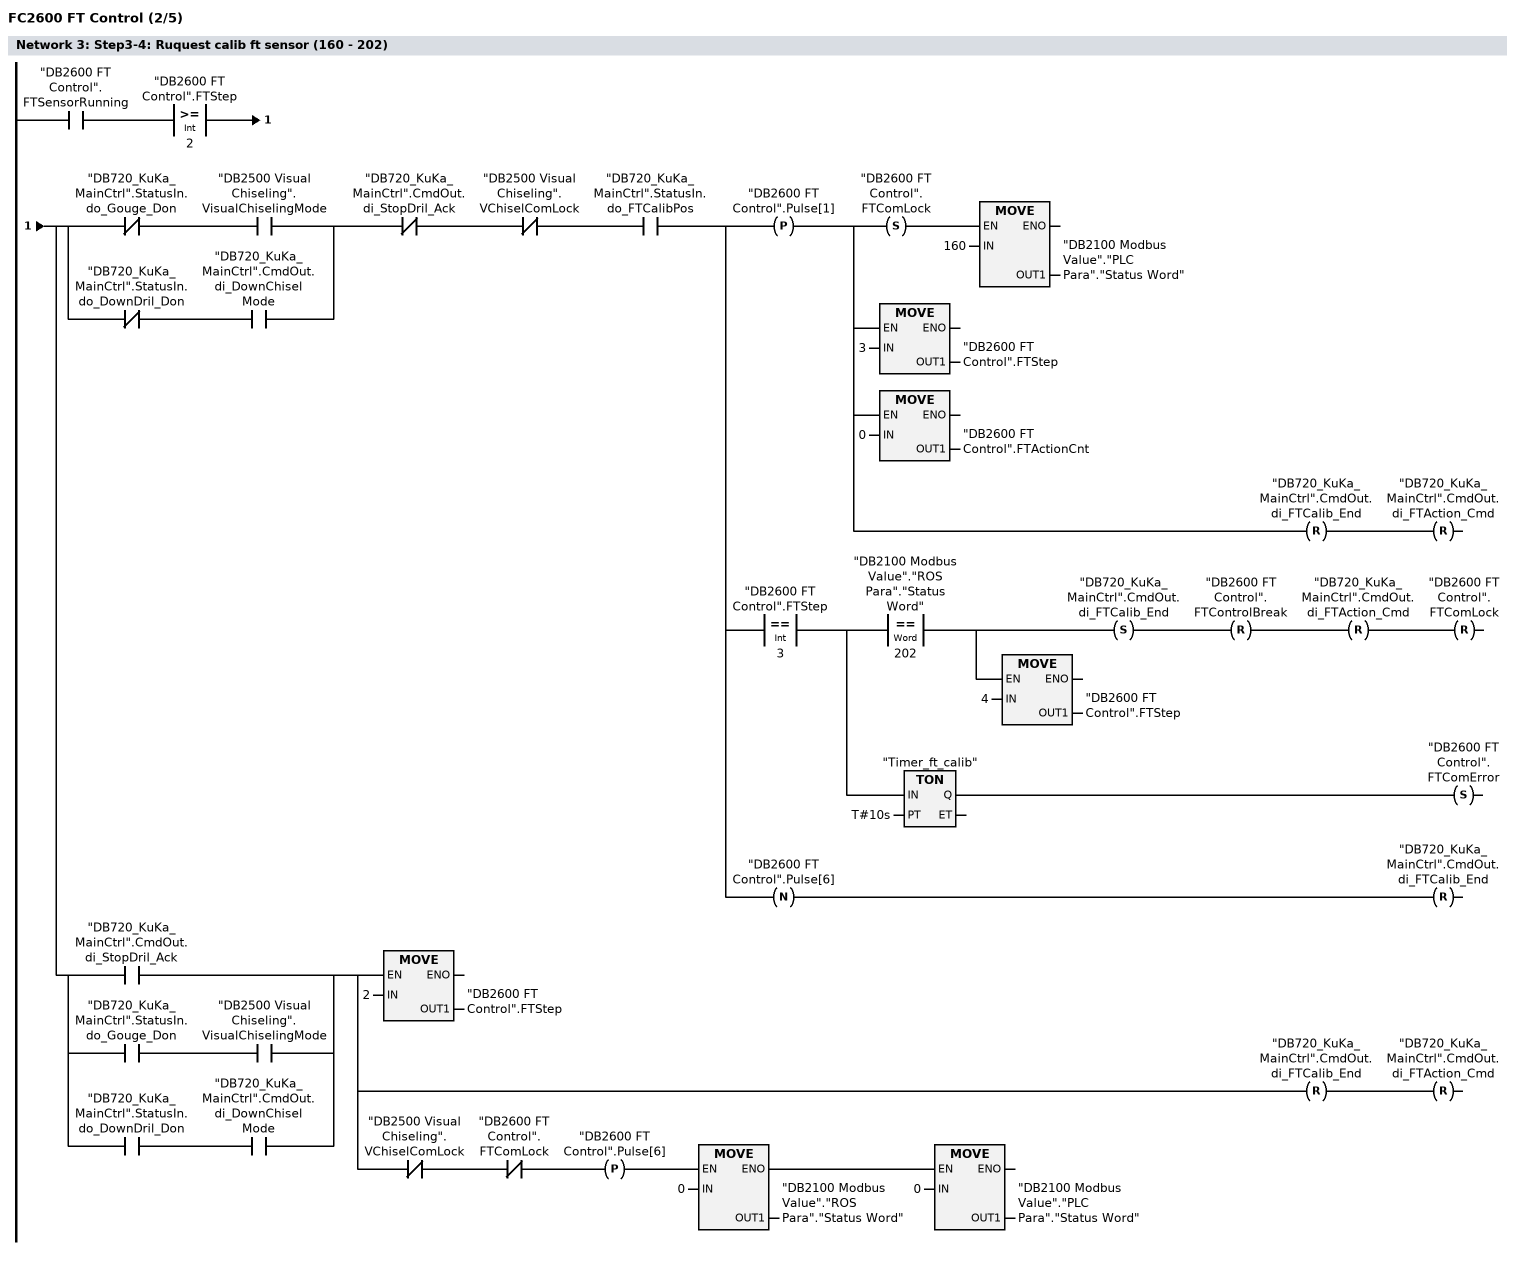
   #_w1 := "DB2600 FT Control".FTSensorRunning AND ("DB2600 FT Control".FTStep >= 2);
   #_w2 := #_w1 AND ((NOT "DB720_KuKa_MainCtrl".StatusIn.do_Gouge_Don AND "DB2500 Visual Chiseling".VisualChiselingMode) OR (NOT "DB720_KuKa_MainCtrl".StatusIn.do_DownDril_Don AND "DB720_KuKa_MainCtrl".CmdOut.di_DownChiselMode)) AND NOT "DB720_KuKa_MainCtrl".CmdOut.di_StopDril_Ack AND NOT "DB2500 Visual Chiseling".VChiselComLock AND "DB720_KuKa_MainCtrl".StatusIn.do_FTCalibPos;
   #_w3 := #_w2 AND NOT "DB2600 FT Control".Pulse[1];   // rising edge
   "DB2600 FT Control".Pulse[1] := #_w2;
   IF #_w3 THEN
       "DB2600 FT Control".FTComLock := TRUE;
       "DB2100 Modbus Value"."PLC Para"."Status Word" := 160;
       "DB2600 FT Control".FTStep := 3;
       "DB2600 FT Control".FTActionCnt := 0;
       "DB720_KuKa_MainCtrl".CmdOut.di_FTCalib_End := FALSE;
       "DB720_KuKa_MainCtrl".CmdOut.di_FTAction_Cmd := FALSE;
   END_IF;
   #_w4 := #_w2 AND ("DB2600 FT Control".FTStep = 3);
   IF #_w4 AND ("DB2100 Modbus Value"."ROS Para"."Status Word" = 202) THEN
       "DB720_KuKa_MainCtrl".CmdOut.di_FTCalib_End := TRUE;
       "DB2600 FT Control".FTControlBreak := FALSE;
       "DB720_KuKa_MainCtrl".CmdOut.di_FTAction_Cmd := FALSE;
       "DB2600 FT Control".FTComLock := FALSE;
       "DB2600 FT Control".FTStep := 4;
   END_IF;
   "Timer_ft_calib".TON(IN := #_w4, PT := T#10s);
   IF "Timer_ft_calib".Q THEN "DB2600 FT Control".FTComError := TRUE; END_IF;
   #_w5 := NOT #_w2 AND "DB2600 FT Control".Pulse[6];   // falling edge
   "DB2600 FT Control".Pulse[6] := #_w2;
   IF #_w5 THEN "DB720_KuKa_MainCtrl".CmdOut.di_FTCalib_End := FALSE; END_IF;
   #_w6 := #_w1 AND ("DB720_KuKa_MainCtrl".CmdOut.di_StopDril_Ack OR ("DB720_KuKa_MainCtrl".StatusIn.do_Gouge_Don AND "DB2500 Visual Chiseling".VisualChiselingMode) OR ("DB720_KuKa_MainCtrl".StatusIn.do_DownDril_Don AND "DB720_KuKa_MainCtrl".CmdOut.di_DownChiselMode));
   IF #_w6 THEN
       "DB2600 FT Control".FTStep := 2;
       "DB720_KuKa_MainCtrl".CmdOut.di_FTCalib_End := FALSE;
       "DB720_KuKa_MainCtrl".CmdOut.di_FTAction_Cmd := FALSE;
   END_IF;
   #_w7 := #_w6 AND NOT "DB2500 Visual Chiseling".VChiselComLock AND NOT "DB2600 FT Control".FTComLock;
   #_w8 := #_w7 AND NOT "DB2600 FT Control".Pulse[6];   // rising edge
   "DB2600 FT Control".Pulse[6] := #_w7;
   IF #_w8 THEN
       "DB2100 Modbus Value"."ROS Para"."Status Word" := 0;
       "DB2100 Modbus Value"."PLC Para"."Status Word" := 0;
   END_IF;
END_REGION

REGION Network 4: Step5-6: request ft control (165 - 203,204,205)
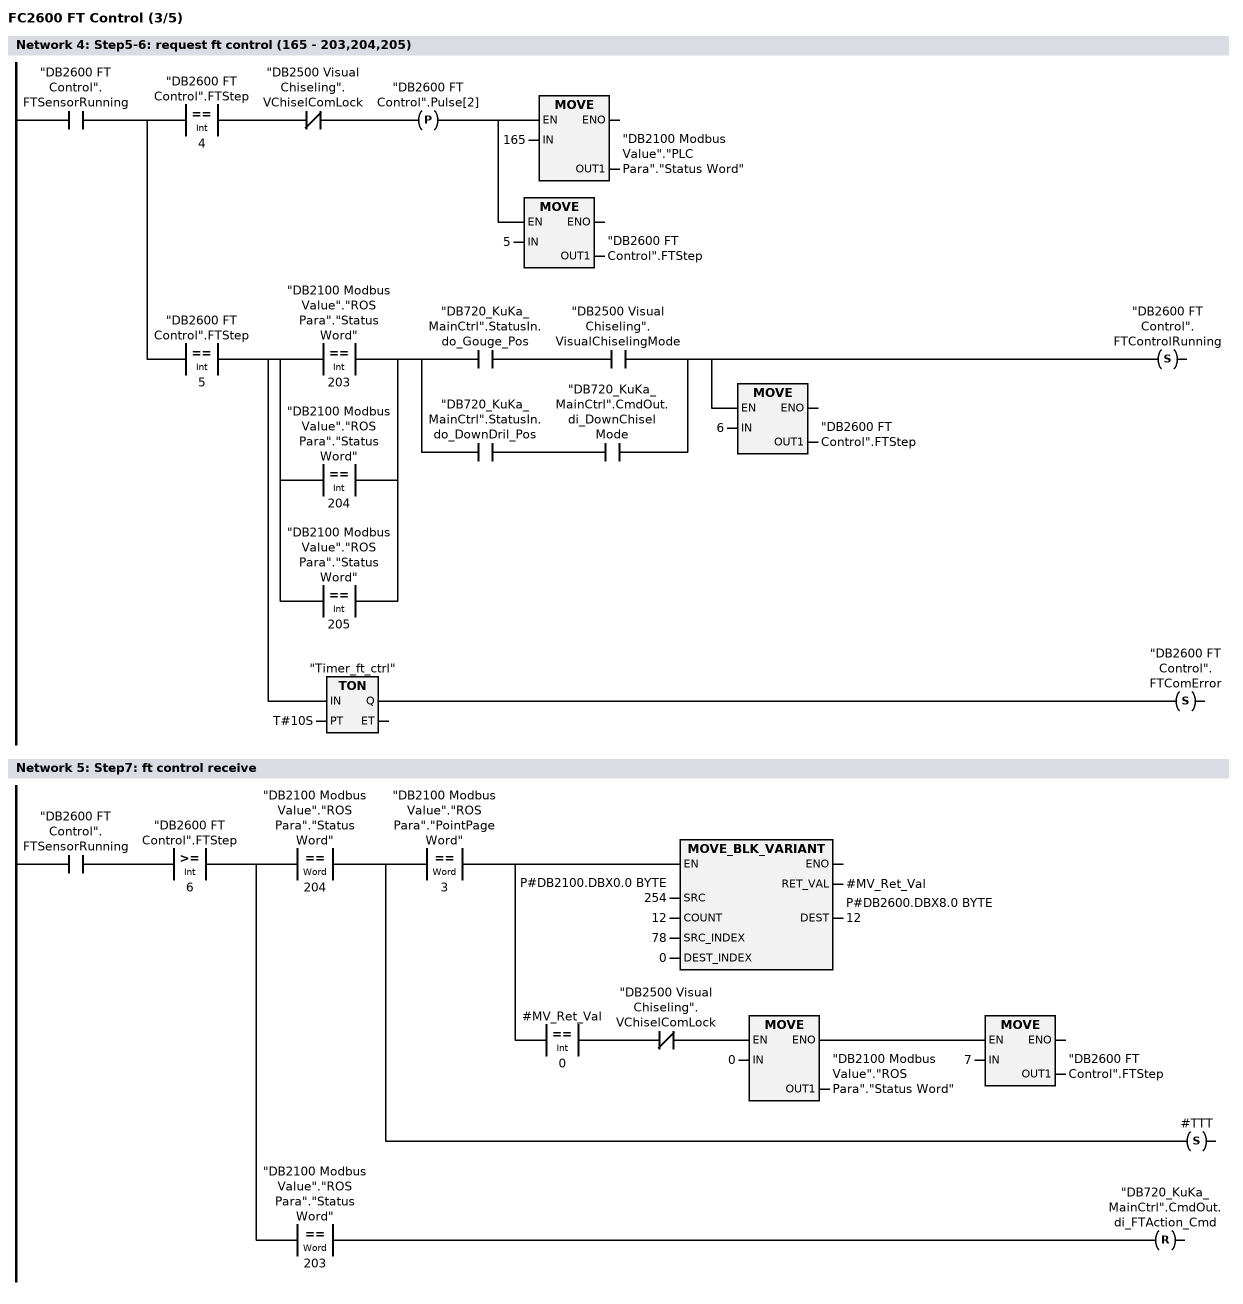
   #_w1 := "DB2600 FT Control".FTSensorRunning AND ("DB2600 FT Control".FTStep = 4) AND NOT "DB2500 Visual Chiseling".VChiselComLock;
   #_w2 := #_w1 AND NOT "DB2600 FT Control".Pulse[2];   // rising edge
   "DB2600 FT Control".Pulse[2] := #_w1;
   IF #_w2 THEN
       "DB2100 Modbus Value"."PLC Para"."Status Word" := 165;
       "DB2600 FT Control".FTStep := 5;
   END_IF;
   #_w3 := "DB2600 FT Control".FTSensorRunning AND ("DB2600 FT Control".FTStep = 5);
   IF #_w3 AND (("DB2100 Modbus Value"."ROS Para"."Status Word" = 203) OR ("DB2100 Modbus Value"."ROS Para"."Status Word" = 204) OR ("DB2100 Modbus Value"."ROS Para"."Status Word" = 205)) AND (("DB720_KuKa_MainCtrl".StatusIn.do_Gouge_Pos AND "DB2500 Visual Chiseling".VisualChiselingMode) OR ("DB720_KuKa_MainCtrl".StatusIn.do_DownDril_Pos AND "DB720_KuKa_MainCtrl".CmdOut.di_DownChiselMode)) THEN
       "DB2600 FT Control".FTControlRunning := TRUE;
       "DB2600 FT Control".FTStep := 6;
   END_IF;
   "Timer_ft_ctrl".TON(IN := #_w3, PT := T#10S);
   IF "Timer_ft_ctrl".Q THEN "DB2600 FT Control".FTComError := TRUE; END_IF;
END_REGION

REGION Network 5: Step7: ft control receive
   #_w1 := "DB2600 FT Control".FTSensorRunning AND ("DB2600 FT Control".FTStep >= 6);
   #_w2 := #_w1 AND ("DB2100 Modbus Value"."ROS Para"."Status Word" = 204);
   #_w3 := #_w2 AND ("DB2100 Modbus Value"."ROS Para"."PointPage Word" = 3);
   IF #_w3 THEN
       #MV_Ret_Val := MOVE_BLK_VARIANT(SRC := P#DB2100.DBX0.0 BYTE 254,
                               COUNT := 12,
                               SRC_INDEX := 78,
                               DEST_INDEX := 0,
                               DEST => P#DB2600.DBX8.0 BYTE 12);
   END_IF;
   IF #_w3 AND (#MV_Ret_Val = 0) AND NOT "DB2500 Visual Chiseling".VChiselComLock THEN
       "DB2100 Modbus Value"."ROS Para"."Status Word" := 0;
       "DB2600 FT Control".FTStep := 7;
   END_IF;
   IF #_w2 THEN #TTT := TRUE; END_IF;
   IF #_w1 AND ("DB2100 Modbus Value"."ROS Para"."Status Word" = 203) THEN
       "DB720_KuKa_MainCtrl".CmdOut.di_FTAction_Cmd := FALSE;
   END_IF;
END_REGION

REGION Network 6: Step8: ft control convert
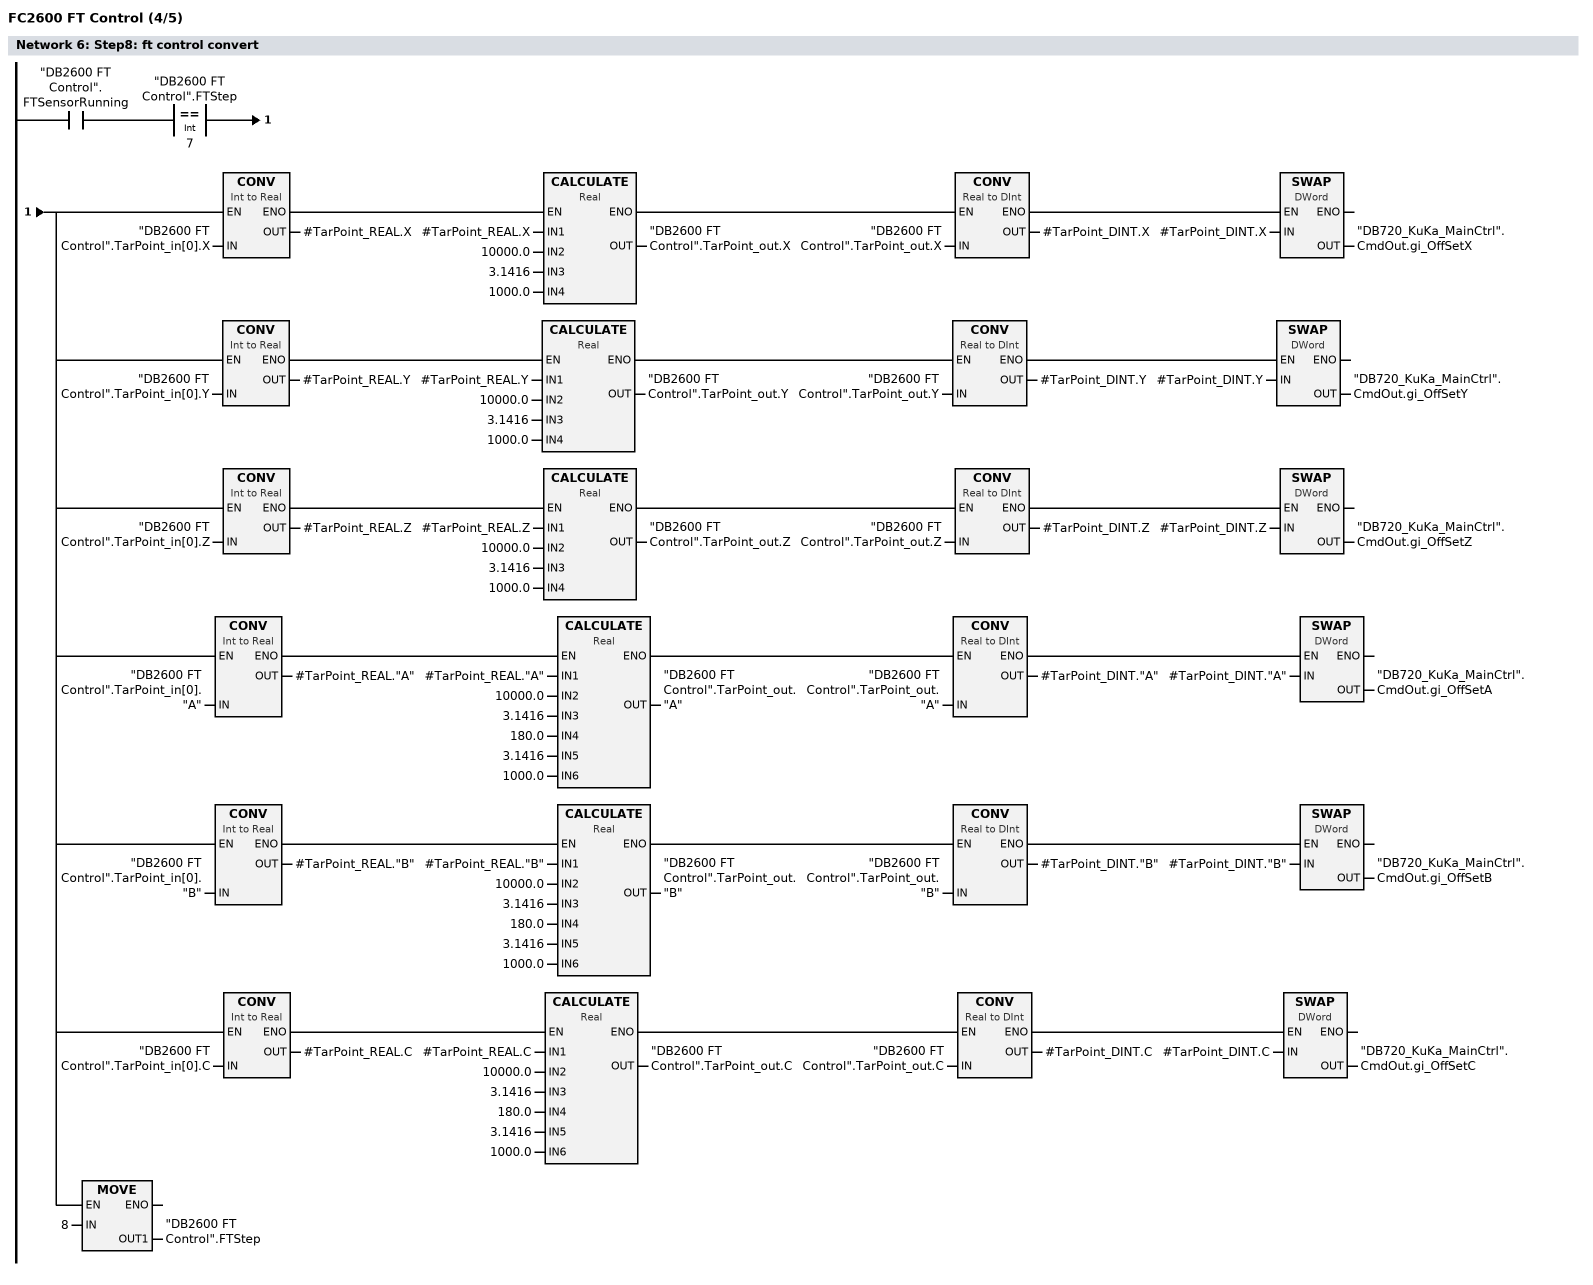
   IF "DB2600 FT Control".FTSensorRunning AND ("DB2600 FT Control".FTStep = 7) THEN
       #TarPoint_REAL.X := INT_TO_REAL("DB2600 FT Control".TarPoint_in[0].X);
       "DB2600 FT Control".TarPoint_out.X := ( #TarPoint_REAL.X / 10000.0 - 3.1416 ) * 1000.0;
       #TarPoint_DINT.X := REAL_TO_DINT("DB2600 FT Control".TarPoint_out.X);
       "DB720_KuKa_MainCtrl".CmdOut.gi_OffSetX := SWAP(#TarPoint_DINT.X);
       #TarPoint_REAL.Y := INT_TO_REAL("DB2600 FT Control".TarPoint_in[0].Y);
       "DB2600 FT Control".TarPoint_out.Y := ( #TarPoint_REAL.Y / 10000.0 - 3.1416 ) * 1000.0;
       #TarPoint_DINT.Y := REAL_TO_DINT("DB2600 FT Control".TarPoint_out.Y);
       "DB720_KuKa_MainCtrl".CmdOut.gi_OffSetY := SWAP(#TarPoint_DINT.Y);
       #TarPoint_REAL.Z := INT_TO_REAL("DB2600 FT Control".TarPoint_in[0].Z);
       "DB2600 FT Control".TarPoint_out.Z := ( #TarPoint_REAL.Z / 10000.0 - 3.1416 ) * 1000.0;
       #TarPoint_DINT.Z := REAL_TO_DINT("DB2600 FT Control".TarPoint_out.Z);
       "DB720_KuKa_MainCtrl".CmdOut.gi_OffSetZ := SWAP(#TarPoint_DINT.Z);
       #TarPoint_REAL."A" := INT_TO_REAL("DB2600 FT Control".TarPoint_in[0]."A");
       "DB2600 FT Control".TarPoint_out."A" := ( ( #TarPoint_REAL."A" / 10000.0 - 3.1416 ) * 180.0 ) / 3.1416*1000.0;
       #TarPoint_DINT."A" := REAL_TO_DINT("DB2600 FT Control".TarPoint_out."A");
       "DB720_KuKa_MainCtrl".CmdOut.gi_OffSetA := SWAP(#TarPoint_DINT."A");
       #TarPoint_REAL."B" := INT_TO_REAL("DB2600 FT Control".TarPoint_in[0]."B");
       "DB2600 FT Control".TarPoint_out."B" := ( ( #TarPoint_REAL."B" / 10000.0 - 3.1416 ) * 180.0 ) / 3.1416*1000.0;
       #TarPoint_DINT."B" := REAL_TO_DINT("DB2600 FT Control".TarPoint_out."B");
       "DB720_KuKa_MainCtrl".CmdOut.gi_OffSetB := SWAP(#TarPoint_DINT."B");
       #TarPoint_REAL.C := INT_TO_REAL("DB2600 FT Control".TarPoint_in[0].C);
       "DB2600 FT Control".TarPoint_out.C := ( ( #TarPoint_REAL.C / 10000.0 - 3.1416 ) * 180.0 ) / 3.1416*1000.0;
       #TarPoint_DINT.C := REAL_TO_DINT("DB2600 FT Control".TarPoint_out.C);
       "DB720_KuKa_MainCtrl".CmdOut.gi_OffSetC := SWAP(#TarPoint_DINT.C);
       "DB2600 FT Control".FTStep := 8;
   END_IF;
END_REGION

REGION Network 7: Step9: ft control send
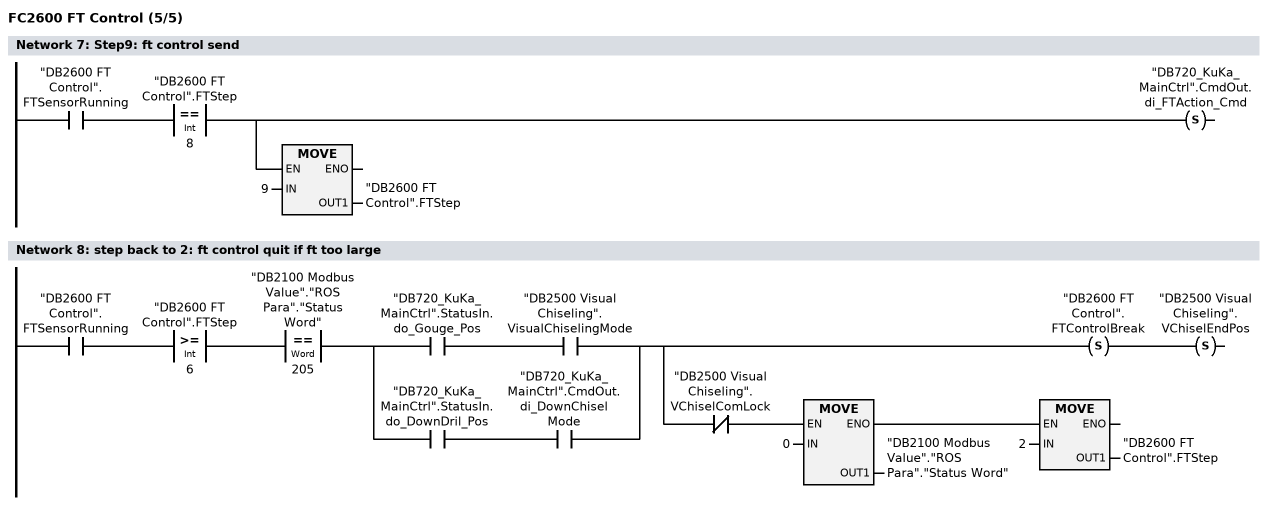
   RUNG wire#powerrail
      Contact( "DB2600 FT Control".FTSensorRunning )
      { S7_Templates := "SrcType := Int" } EQ_Contact(in1 := "DB2600 FT Control".FTStep, in2 := 8)
      wire#w1
      S_Coil( "DB720_KuKa_MainCtrl".CmdOut.di_FTAction_Cmd )
   END_RUNG
   RUNG wire#w1
      Move(in := 9, out1 => "DB2600 FT Control".FTStep)
   END_RUNG
   // the same network as SCL:
   IF "DB2600 FT Control".FTSensorRunning AND ("DB2600 FT Control".FTStep = 8) THEN
       "DB720_KuKa_MainCtrl".CmdOut.di_FTAction_Cmd := TRUE;
       "DB2600 FT Control".FTStep := 9;
   END_IF;
END_REGION

REGION Network 8: step back to 2: ft control quit if ft too large
   RUNG wire#powerrail
      Contact( "DB2600 FT Control".FTSensorRunning )
      { S7_Templates := "SrcType := Int" } GE_Contact(in1 := "DB2600 FT Control".FTStep, in2 := 6)
      { S7_Templates := "SrcType := Word" } EQ_Contact(in1 := "DB2100 Modbus Value"."ROS Para"."Status Word", in2 := 205)
      wire#w1
      Contact( "DB720_KuKa_MainCtrl".StatusIn.do_Gouge_Pos )
      Contact( "DB2500 Visual Chiseling".VisualChiselingMode )
      wire#w2
      S_Coil( "DB2600 FT Control".FTControlBreak )
      S_Coil( "DB2500 Visual Chiseling".VChiselEndPos )
   END_RUNG
   RUNG wire#w1
      Contact( "DB720_KuKa_MainCtrl".StatusIn.do_DownDril_Pos )
      Contact( "DB720_KuKa_MainCtrl".CmdOut.di_DownChiselMode )
   END_RUNG wire#w2
   RUNG wire#w2
      I_Contact( "DB2500 Visual Chiseling".VChiselComLock )
      Move(in := 0, out1 => "DB2100 Modbus Value"."ROS Para"."Status Word")
      Move(in := 2, out1 => "DB2600 FT Control".FTStep)
   END_RUNG
   // the same network as SCL:
   #_w1 := "DB2600 FT Control".FTSensorRunning AND ("DB2600 FT Control".FTStep >= 6) AND ("DB2100 Modbus Value"."ROS Para"."Status Word" = 205) AND (("DB720_KuKa_MainCtrl".StatusIn.do_Gouge_Pos AND "DB2500 Visual Chiseling".VisualChiselingMode) OR ("DB720_KuKa_MainCtrl".StatusIn.do_DownDril_Pos AND "DB720_KuKa_MainCtrl".CmdOut.di_DownChiselMode));
   IF #_w1 THEN
       "DB2600 FT Control".FTControlBreak := TRUE;
       "DB2500 Visual Chiseling".VChiselEndPos := TRUE;
   END_IF;
   IF #_w1 AND NOT "DB2500 Visual Chiseling".VChiselComLock THEN
       "DB2100 Modbus Value"."ROS Para"."Status Word" := 0;
       "DB2600 FT Control".FTStep := 2;
   END_IF;
END_REGION
END_FUNCTION

// folder: 099_systemErrOB

ORGANIZATION_BLOCK "Pull or plug of modules"   // OB83, LAD, PullPlug
{ S7_Optimized_Access := 'TRUE' }
VERSION : 0.1
   VAR_INPUT
      LADDR : Hw_Io;   // Hardware identifier
      Event_Class : Byte;   // 16#38/39: module inserted, removed
      Fault_ID : Byte;   // Fault identifier
   END_VAR
BEGIN
END_ORGANIZATION_BLOCK

ORGANIZATION_BLOCK "Rack or station failure"   // OB86, LAD, RackStationFailure
{ S7_Optimized_Access := 'TRUE' }
VERSION : 0.1
   VAR_INPUT
      LADDR : Hw_Io;   // Hardware identifier
      Event_Class : Byte;   // Event class
      Fault_ID : Byte;   // Fault identifier
   END_VAR
BEGIN
END_ORGANIZATION_BLOCK

ORGANIZATION_BLOCK "Startup"   // OB100, LAD, Startup
TITLE = "Complete Restart"
{ S7_Optimized_Access := 'TRUE' }
VERSION : 0.1
   VAR_INPUT
      LostRetentive : Bool;   // True if retentive data are lost
      LostRTC : Bool;   // True if date and time are lost
   END_VAR
BEGIN
END_ORGANIZATION_BLOCK

ORGANIZATION_BLOCK "System Err"   // OB123, LAD, ProgramCycle
TITLE = "Main Program Sweep (Cycle)"
{ S7_Optimized_Access := 'TRUE' }
VERSION : 0.1
   VAR_INPUT
      Initial_Call : Bool;   // Initial call of this OB
      Remanence : Bool;   // =True, if remanent data are available
   END_VAR
BEGIN
END_ORGANIZATION_BLOCK

(* ===== HMI "HMI_RT_1" =====

ScreenModuleEditorView "Faceplate_1" 640x480
   TextField "文本域_7" at 221,13 size 76x20; Text '设定速度: / 当前速度'
   TextField "文本域_9" at 217,13 size 108x20; Text '扭矩目标/Nm： / 当前速度'
   TextField "文本域_13" at 446,15 size 84x20; Text '位置表编号 / 当前速度'
   TextField "文本域_8" at 221,83 size 76x20; Text '设定速度: / 当前速度'
   TextField "文本域_15" at 211,81 size 100x20; Text '读出参数值： / 当前速度'
   TextField "文本域_19" at 330,81 size 100x20; Text '写入参数值： / 当前速度'
   TextField "文本域_17" at 211,52 size 116x20; Text '通讯参数编号： / 当前速度'
   IOField "IO 域_2" at 327,10 size 116x31; FormatPattern 999.99
   Button "按钮_12" at 10,10 size 200x64; TextOff '电机扭矩模式 启动 ST02伺服 点动前进'; TextList "Cylinder_Name_1"
   Button "按钮_2" at 529,10 size 116x64; TextOff '位置表 启动 ST02伺服 点动前进'; TextList "Cylinder_Name_1"
   IOField "IO 域_3" at 445,42 size 83x32; FormatPattern 99
   Button "按钮_7" at 10,76 size 200x64; TextOff '读取参数 ST02伺服 点动前进'; TextList "Cylinder_Name_1"
   IOField "IO 域_5" at 327,43 size 116x31; FormatPattern 999999
   IOField "IO 域_10" at 212,107 size 115x33; FormatPattern 99999999.99
   Button "按钮_6" at 445,76 size 200x64; TextOff '写入参数 ST02伺服 点动前进'; TextList "Cylinder_Name_1"
   IOField "IO 域_4" at 328,107 size 115x33; FormatPattern 99999999.99
*)

(* ===== HMI "HMI_RT_1" =====

ScreenModuleEditorView "Faceplate_1" 640x480
   TextField "文本域_7" at 221,13 size 76x20; Text '设定速度: / 当前速度'
   TextField "文本域_9" at 217,13 size 108x20; Text '扭矩目标/Nm： / 当前速度'
   TextField "文本域_13" at 446,15 size 84x20; Text '位置表编号 / 当前速度'
   TextField "文本域_8" at 221,83 size 76x20; Text '设定速度: / 当前速度'
   TextField "文本域_15" at 211,81 size 100x20; Text '读出参数值： / 当前速度'
   TextField "文本域_19" at 330,81 size 100x20; Text '写入参数值： / 当前速度'
   TextField "文本域_17" at 211,52 size 116x20; Text '通讯参数编号： / 当前速度'
   IOField "IO 域_2" at 327,10 size 116x31; FormatPattern 999.99
   Button "按钮_12" at 10,10 size 200x64; TextOff '电机扭矩模式 启动 ST02伺服 点动前进'; TextList "Cylinder_Name_1"
   Button "按钮_2" at 529,10 size 116x64; TextOff '位置表 启动 ST02伺服 点动前进'; TextList "Cylinder_Name_1"
   IOField "IO 域_3" at 445,42 size 83x32; FormatPattern 99
   Button "按钮_7" at 10,76 size 200x64; TextOff '读取参数 ST02伺服 点动前进'; TextList "Cylinder_Name_1"
   IOField "IO 域_5" at 327,43 size 116x31; FormatPattern 999999
   IOField "IO 域_10" at 212,107 size 115x33; FormatPattern 99999999.99
   Button "按钮_6" at 445,76 size 200x64; TextOff '写入参数 ST02伺服 点动前进'; TextList "Cylinder_Name_1"
   IOField "IO 域_4" at 328,107 size 115x33; FormatPattern 99999999.99
*)

(* ===== HMI "HMI_RT_1" =====
system functions are stored by id; their names below are inferred from use
connection "PLC_1200": ETHERNET, S7_1200_OMS

HMI tags "默认变量表"
   "Language" : Int, internal
   "DB_Message_PromptValue" : Int = PLC DB1140_Message.PromptValue, 1 s
   "Page" : Int, internal
   "SerialCom_Index" : Int, internal
   "DB_AutoStep_CycleTime_CycleTime_Net" : Time = PLC DB1060_AutoStep.CycleTime.CycleTime_Net, 1 s
   "DB_Parameter_TypeParaE_Other_FixtureEnable" : Bool = PLC DB1010_Parameter.TypeParaE.Other.FixtureEnable AT %DB1010.DBX922.0, 1 s
   "DB_ValveCall_ST01_Z02_RetPos" : Bool = PLC DB1081_ValveCall.ST01.Z02.RetPos AT %DB1081.DBX7.3, 1 s
   "DB_ValveCall_ST01_Z02_ExtPos" : Bool = PLC DB1081_ValveCall.ST01.Z02.ExtPos AT %DB1081.DBX7.2, 1 s
   "DB_ValveCall_ST01_Z02_ExtPmt" : Bool = PLC DB1081_ValveCall.ST01.Z02.ExtPmt AT %DB1081.DBX6.2, 1 s
   "DB_ValveCall_ST01_Z02_RetPmt" : Bool = PLC DB1081_ValveCall.ST01.Z02.RetPmt AT %DB1081.DBX6.3, 1 s
   "DB_ValveCall_ST01_Z02_RetTPPB" : Bool = PLC DB1081_ValveCall.ST01.Z02.RetTPPB AT %DB1081.DBX6.1, 1 s
   "DB_ValveCall_ST01_Z02_ExtTPPB" : Bool = PLC DB1081_ValveCall.ST01.Z02.ExtTPPB AT %DB1081.DBX6.0, 1 s
   "DB_Timer_Communication" : Bool = PLC DB1042_Timer.Communication AT %DB1042.DBX0.0, 1 s
   "DB_Component_Analog_Out_Ctrl_IN_Target" : Real = PLC DB1080_Component.Analog_Out_1.Ctrl_Out.Pressure AT %DB1080.DBD474, 1 s
   "DB_Component_Aux_Pressure" : Real = PLC DB1080_Component.Aux.Pressure AT %DB1080.DBD938, 1 s
   "DB_KuKa_MainCtrl.Aux.CheckNo" : Int = PLC DB720_KuKa_MainCtrl.Aux.CheckNo AT %DB720.DBW270, 1 s
   "DB_Timer_Force" : Real = PLC DB1042_Timer.Force AT %DB1042.DBD14, 1 s

HMI tags "System_Para"
   "DB_Component_Aux_SysTimeSet_YEAR" : UInt = PLC DB1080_Component.Aux.SysTimeSet.YEAR AT %DB1080.DBW970, 1 s
   "DB_Component_Aux_SysTimeSet_MONTH" : USInt = PLC DB1080_Component.Aux.SysTimeSet.MONTH AT %DB1080.DBB972, 1 s

HMI tags "DB_Parameter_Base"
   "DB_Parameter_TP_Cmd" : Word = PLC DB1010_Parameter.TP_Cmd, 1 s
   "DB_Parameter_AryTypeName(9)" : String[20] = PLC DB1010_Parameter.AryTypeName[9], 1 s   // 产品型号选择页面显示的产品名称；
   "DB_Parameter_AryTypeName(2)" : String[20] = PLC DB1010_Parameter.AryTypeName[2], 1 s   // 产品型号选择页面显示的产品名称；
   "DB_Parameter_AryTypeName(11)" : String[20] = PLC DB1010_Parameter.AryTypeName[11], 1 s   // 产品型号选择页面显示的产品名称；
   "DB_Parameter_AryTypeName(3)" : String[20] = PLC DB1010_Parameter.AryTypeName[3], 1 s   // 产品型号选择页面显示的产品名称；
   "DB_Parameter_AryTypeName(5)" : String[20] = PLC DB1010_Parameter.AryTypeName[5], 1 s   // 产品型号选择页面显示的产品名称；
   "DB_Parameter_AryTypeName(4)" : String[20] = PLC DB1010_Parameter.AryTypeName[4], 1 s   // 产品型号选择页面显示的产品名称；
   "DB_Parameter_TypeParaR_TypeName" : String[20] = PLC DB1010_Parameter.TypeParaR.TypeName, 1 s
   "DB_Parameter_AryTypeName(8)" : String[20] = PLC DB1010_Parameter.AryTypeName[8], 1 s   // 产品型号选择页面显示的产品名称；
   "DB_Parameter_TypeParaE_TypeName" : String[20] = PLC DB1010_Parameter.TypeParaE.TypeName, 1 s
   "DB_Parameter_AryTypeName(1)" : String[20] = PLC DB1010_Parameter.AryTypeName[1], 1 s   // 产品型号选择页面显示的产品名称；
   "DB_Parameter_AryTypeName(7)" : String[20] = PLC DB1010_Parameter.AryTypeName[7], 1 s   // 产品型号选择页面显示的产品名称；
   "DB_Parameter_AryTypeName(6)" : String[20] = PLC DB1010_Parameter.AryTypeName[6], 1 s   // 产品型号选择页面显示的产品名称；
   "DB_Parameter_CurProgNoE" : Int = PLC DB1010_Parameter.CurProgNoE, 1 s   // 当前程序号编辑区；
   "DB_Parameter_TP_Status" : Word = PLC DB1010_Parameter.TP_Status, 1 s
   "DB_Parameter_ArrayProgNoForSel" : Array [0..9] of Int = PLC DB1010_Parameter.ArrayProgNoForSel, 1 s
   "DB_Parameter_AryTypeName(10)" : String[20] = PLC DB1010_Parameter.AryTypeName[10], 1 s
   "DB_Parameter_CurProgNoR" : Int = PLC DB1010_Parameter.CurProgNoR, 1 s
   "DB_Parameter_ProgNoCopyDest" : Int = PLC DB1010_Parameter.ProgNoCopyDest, 1 s
   "DB_Parameter_IMaxProgNo" : Int = PLC DB1010_Parameter.IMaxProgNo, 1 s

HMI tags "Standard_Switch"
   "Cylinder_Index_Max" : Int, internal   // 到达最大气缸数
   "Cylinder_Index_Min" : Int, internal   // 到达最小气缸数
   "手动控制\CylinderIndex1" : Int, internal
   "手动控制\CylinderIndex2" : Int, internal
   "手动控制\CylinderIndex3" : Int, internal
   "手动控制\CylinderIndex4" : Int, internal
   "手动控制\CylinderIndex5" : Int, internal
   "Z01_Cmd" : Byte AT %DB1081.DBB0, 100 ms   // 气缸名1
   "Z02_CmdW" : Byte AT %DB1081.DBB0, 100 ms   // 气缸名1
   "Z03_CmdW" : Byte AT %DB1081.DBB0, 100 ms   // 气缸名1
   "Z04_CmdW" : Byte AT %DB1081.DBB0, 100 ms   // 气缸名1
   "Z05_CmdW" : Byte AT %DB1081.DBB0, 100 ms   // 气缸名1
   "Z01_Status" : Word AT %DB1081.DBW0, 100 ms   // 气缸名1
   "Z02_Status" : Word AT %DB1081.DBW0, 100 ms   // 气缸名1
   "Z03_Status" : Word AT %DB1081.DBW0, 100 ms   // 气缸名1
   "Z04_Status" : Word AT %DB1081.DBW0, 100 ms   // 气缸名1
   "Z05_Status" : Word AT %DB1081.DBW0, 100 ms   // 气缸名1
   "Cyl_Addr_Z01" : UInt, internal
   "Cyl_Addr_Z02" : UInt, internal
   "Cyl_Addr_Z03" : UInt, internal
   "Cyl_Addr_Z04" : UInt, internal
   "Cyl_Addr_Z05" : UInt, internal
   "DB_SysMode_Cylinder_Index" : Int = PLC DB1001_SysMode.Cylinder_Index, 100 ms   // 触摸屏中选择的气缸编号,从1计数
      on ChangeValue: function_dbe01993("手动控制\CylinderIndex1", 1, "DB_SysMode_Cylinder_Index", 0); function_dbe01993("手动控制\CylinderIndex2", 1, "DB_SysMode_Cylinder_Index", 1); function_dbe01993("手动控制\CylinderIndex3", 1, "DB_SysMode_Cylinder_Index", 2); function_dbe01993("手动控制\CylinderIndex4", 1, "DB_SysMode_Cylinder_Index", 3); function_dbe01993("手动控制\CylinderIndex5", 1, "DB_SysMode_Cylinder_Index", 4); function_dbe01993("Cyl_Addr_Z01", 6, "DB_SysMode_Cylinder_Index", -6); function_dbe01993("Cyl_Addr_Z02", 6, "DB_SysMode_Cylinder_Index", 0); function_dbe01993("Cyl_Addr_Z03", 6, "DB_SysMode_Cylinder_Index", 6); function_dbe01993("Cyl_Addr_Z04", 6, "DB_SysMode_Cylinder_Index", 12); function_dbe01993("Cyl_Addr_Z05", 6, "DB_SysMode_Cylinder_Index", 18)

HMI tags "DB_Err"
   "Err009" : Word AT %DB1148.DBW16, 1 s
   "Err008" : Word AT %DB1148.DBW14, 1 s
   "Err007" : Word AT %DB1148.DBW12, 1 s
   "Err006" : Word AT %DB1148.DBW10, 1 s
   "Err005" : Word AT %DB1148.DBW8, 1 s
   "Err004" : Word AT %DB1148.DBW6, 1 s
   "Err003" : Word AT %DB1148.DBW4, 1 s
   "Err002" : Word AT %DB1148.DBW2, 1 s
   "Err012" : Word AT %DB1148.DBW22, 1 s
   "Err011" : Word AT %DB1148.DBW20, 1 s
   "Err010" : Word AT %DB1148.DBW18, 1 s
   "Err001" : Word AT %DB1148.DBW0, 1 s
   "Err013" : Word AT %DB1148.DBW24, 1 s
   "Err014" : Word AT %DB1148.DBW26, 1 s
   "Err015" : Word AT %DB1148.DBW28, 1 s
   "Err016" : Word AT %DB1148.DBW30, 1 s
   "Err017" : Word AT %DB1148.DBW32, 1 s
   "Err018" : Word AT %DB1148.DBW34, 1 s
   "Err019" : Word AT %DB1148.DBW36, 1 s
   "Err020" : Word AT %DB1148.DBW38, 1 s
   "Err021" : Word AT %DB1148.DBW40, 1 s
   "Err022" : Word AT %DB1148.DBW42, 1 s

HMI tags "Addr_DB_SysMode"
   "Addr_DB_SysMode_Mode" : Int, internal
   "Addr_DB_SysMode_TPCurPageType" : Int, internal
   "Addr_DB_SysMode_TPCurSubPage" : Int, internal
   "Addr_DB_SysMode_TPPB" : Int, internal
   "Addr_DB_SysMode_TPSetPageNO" : Int, internal
   "Addr_DB_SysMode_Status" : Int, internal
   "Addr_DB_SysMode_IO_FromTP" : Int, internal
   "Addr_DB_SysMode_IO_Cur" : Int, internal
   "Addr_DB_SysMode_Output" : Int, internal

HMI tags "DB_Sys_Public"
   "DB_SysMode_Sys_Time_CurPLCTime" : DTL = PLC DB1001_SysMode.Sys_Time.CurPLCTime, 1 s
   "DB_SysMode_Sys_Time_SetPLCTimeTP" : DTL = PLC DB1001_SysMode.Sys_Time.SetPLCTimeTP, 1 s
   "DB_SysMode_TP_Cmd" : Word = PLC DB1001_SysMode.TP_Cmd, 1 s
   "DB_SysMode_SysMode_Station_Index" : Int = PLC DB1001_SysMode.SysMode_Station_Index, 1 s
      on ChangeValue: function_dbe01993("Addr_DB_SysMode_Mode", 200, "DB_SysMode_SysMode_Station_Index", 10); function_dbe01993("Addr_DB_SysMode_TPPB", 200, "DB_SysMode_SysMode_Station_Index", 18); function_dbe01993("Addr_DB_SysMode_Status", 200, "DB_SysMode_SysMode_Station_Index", 24); function_dbe01993("Addr_DB_SysMode_TPSetPageNO", 200, "DB_SysMode_SysMode_Station_Index", 26); function_dbe01993("Addr_DB_SysMode_TPCurPageType", 200, "DB_SysMode_SysMode_Station_Index", 28); function_dbe01993("Addr_DB_SysMode_TPCurSubPage", 200, "DB_SysMode_SysMode_Station_Index", 30); function_dbe01993("Addr_DB_SysMode_IO_FromTP", 200, "DB_SysMode_SysMode_Station_Index", 32); function_dbe01993("Addr_DB_SysMode_IO_Cur", 200, "DB_SysMode_SysMode_Station_Index", 34); function_dbe01993("Addr_DB_SysMode_Output", 200, "DB_SysMode_SysMode_Station_Index", 4)
   "DB_SysMode_DisableOption" : Word AT %DB1001.DBW0, 1 s

HMI tags "DB_SysMode"
   "DB_SysMode_TPSetPageNo" : Int AT %DB1001.DBW0, 500 ms
      on ChangeValue: ActivateScreenByNumber("DB_SysMode_TPSetPageNo", 1)
   "DB_SysMode_TPCurSubPage" : Int AT %DB1001.DBW0, 1 s
   "DB_SysMode_TPCurPageType" : Int AT %DB1001.DBW0, 1 s
   "DB_SysMode_TPPB" : Word AT %DB1001.DBW0, 1 s
   "DB_SysMode_ModeByte" : Byte AT %DB1001.DBB0, 1 s   // Byte类型的模式开关
   "DB_SysMode_Status" : Word AT %DB1001.DBW0, 100 ms
   "DB_SysMode_IO_FromTP" : Int AT %DB1001.DBW0, 1 s
   "DB_SysMode_IO_Cur" : Int AT %DB1001.DBW0, 1 s
   "DB_SysMode_IO_FromTP_BitArray" : Array [0..15] of Bool AT %DB1001.DBX0.0, 1 s
   "DB_SysMode_Output" : Word AT %DB1001.DBW0, 100 ms
   "DB_SysMode_TPPB_BitArray" : Array [0..15] of Bool AT %DB1001.DBX0.0, 1 s

HMI tags "IO_Check"
   "DB_IOCheck____In_ByteNo" : Int = PLC DB1202_IOCheck.In_ByteNo, 1 s   // Out当前要显示的Byte编号IB0，ByteNo=0
   "DB_IOCheck____In_ByteNo_X10" : Array [0..7] of Int = PLC DB1202_IOCheck.In_ByteNo_X10, 1 s   // 用于更新当前显示Input的内容；
   "IO_Input_SignalStatus" : Byte AT %IB0, 1 s   // 当前显示InPut的On_Off状态信息
   "DB_IOCheck____InputMaxByteNo" : Int = PLC DB1202_IOCheck.InputMaxByteNo, 1 s   // 输入IO最大Byte地址
   "DB_IOCheck____InputMinByteNo" : Int = PLC DB1202_IOCheck.InputMinByteNo, 1 s   // 输入IO最小Byte地址
   "DB_IOCheck____TP_Status" : Word = PLC DB1202_IOCheck.TP_Status, 1 s   // 上页
   "DB_IOCheck____Out_ByteNo" : Int = PLC DB1202_IOCheck.Out_ByteNo, 1 s   // Out当前要显示的Byte编号IB0，ByteNo=0
   "IO_OutPut_SignalStatus" : Byte AT %QB0, 1 s   // 当前显示OutPut的On_Off状态信息
   "DB_IOCheck____OutputMaxByteNo" : Int = PLC DB1202_IOCheck.OutputMaxByteNo, 1 s   // 输出IO最大Byte地址
   "DB_IOCheck____OutputMinByteNo" : Int = PLC DB1202_IOCheck.OutputMinByteNo, 1 s   // 输出IO最小Byte地址
   "DB_IOCheck____Out_ByteNo_X10" : Array [0..7] of Int = PLC DB1202_IOCheck.Out_ByteNo_X10, 1 s

HMI tags "Component_Public"
   "ObjectComment" : WString[80], internal
   "Unit_Position" : WString[10], internal
   "Unit_Speed" : WString[10], internal
   "Unit_Analog" : WString[10], internal
   "Unit_LeakRate" : WString[10], internal
   "Unit_LeakTestPressure" : WString[10], internal
   "Object_Description" : WString[100], internal

HMI tags "KuKaRobot"
   "DB_Component_Robot_TP_Cmd" : Word = PLC DB1080_Component.Robot.TP_Cmd AT %DB1080.DBW2, 1 s
   "DB_Component_Robot_TP_Status" : Word = PLC DB1080_Component.Robot.TP_Status AT %DB1080.DBW4, 1 s
   "DB_Component_Robot_CTRL_IN_ProgNo" : Byte = PLC DB1080_Component.Robot.CTRL_IN.ProgNo AT %DB1080.DBB8, 1 s
   "DB_Component_Robot_CTRL_OUT_ProgNo" : Byte = PLC DB1080_Component.Robot.CTRL_OUT.ProgNo AT %DB1080.DBB36, 1 s
   "DB_Component_Robot_CTRL_OUT_AppInfNo" : Byte = PLC DB1080_Component.Robot.CTRL_OUT.AppInfNo AT %DB1080.DBB37, 1 s
   "DB_Component_Robot_CTRL_OUT_ErrorCode" : Word = PLC DB1080_Component.Robot.CTRL_OUT.ErrorCode AT %DB1080.DBW38, 1 s
   "DB_Component_Robot_CTRL_OUT_LastCylceTime" : Time = PLC DB1080_Component.Robot.CTRL_OUT.LastCylceTime AT %DB1080.DBD40, 1 s
   "DB_Component_Robot_Step_Main" : Int = PLC DB1080_Component.Robot.Step.Main AT %DB1080.DBW64, 1 s
   "DB_Component_Robot_CTRL_IN_RobotSpeed" : Byte = PLC DB1080_Component.Robot.CTRL_IN.RobotSpeed AT %DB1080.DBB9, 1 s
   "DB_Component_Robot_Status_PromptValue" : Int = PLC DB1080_Component.Robot.Status.PromptValue AT %DB1080.DBW62, 1 s
   "AG1520RobotIndex" : UInt AT %DB1.DBW0
   "DB_KuKa_MainCtrl_Ctrl_In_LoadBoxIndex" : Byte = PLC DB720_KuKa_MainCtrl.Ctrl_In.LoadBoxIndex AT %DB720.DBB113, 1 s
   "DB_KuKa_MainCtrl_Ctrl_In_GearBoxIndex" : Byte = PLC DB720_KuKa_MainCtrl.Ctrl_In.GearBoxIndex AT %DB720.DBB112, 1 s
   "DB_KuKa_MainCtrl_Ctrl_In_ProductIndex" : Byte = PLC DB720_KuKa_MainCtrl.Ctrl_In.ProductIndex AT %DB720.DBB116, 1 s
   "DB_KuKa_MainCtrl_Ctrl_In_AssemblyBoxDirection" : Byte = PLC DB720_KuKa_MainCtrl.Ctrl_In.AssemblyBoxDirection AT %DB720.DBB115, 1 s
   "DB_KuKa_MainCtrl_Ctrl_In_ProductBoxDirection" : Byte = PLC DB720_KuKa_MainCtrl.Ctrl_In.ProductBoxDirection AT %DB720.DBB117, 1 s
   "DB_KuKa_MainCtrl_Ctrl_In_UnloadBoxIndex" : Byte = PLC DB720_KuKa_MainCtrl.Ctrl_In.UnloadBoxIndex AT %DB720.DBB114, 1 s
   "DB_KuKa_MainCtrl.CheckAiguille.StartCmd" : Bool = PLC DB720_KuKa_MainCtrl.CheckBit.StartCmd AT %DB720.DBX116.1, 1 s
   "DB_KuKa_MainCtrl.DrillHorizontal.StartCmd" : Bool = PLC DB1060_AutoStep.HorDrillAutoStep.HorDrillStep.StartCmd, 1 s
   "DB_KuKa_MainCtrl.CleanTool.StartCmd" : Bool = PLC DB_KuKa_MainCtrl.CleanTool.StartCmd AT %DB720.DBX164.1, 1 s
   "DB_KuKa_MainCtrl.ChangeTool.StartCmd" : Bool = PLC DB720_KuKa_MainCtrl.ChangeTool.StartCmd AT %DB720.DBX126.1, 1 s
   "DB_KuKa_MainCtrl.CheckAiguille.StepStart" : Bool = PLC DB720_KuKa_MainCtrl.CheckBit.StepStart AT %DB720.DBX116.4, 1 s
   "DB_KuKa_MainCtrl.DrillHorizontal.StepStart" : Bool = PLC DB1060_AutoStep.HorDrillAutoStep.HorDrillStep.StepStart, 1 s
   "DB_KuKa_MainCtrl.CleanTool.StepStart" : Bool = PLC DB_KuKa_MainCtrl.CleanTool.StepStart AT %DB720.DBX164.4, 1 s
   "DB_KuKa_MainCtrl.ChangeTool.StepStart" : Bool = PLC DB720_KuKa_MainCtrl.ChangeTool.StepStart AT %DB720.DBX126.4, 1 s
   "DB_KuKa_MainCtrl.DrillDownload.StartCmd" : Bool = PLC DB720_KuKa_MainCtrl.DrillDownload.StartCmd AT %DB720.DBX134.1, 1 s
   "DB_KuKa_MainCtrl.DrillUpload.StartCmd" : Bool = PLC DB720_KuKa_MainCtrl.DrillUpload.StartCmd AT %DB720.DBX144.1, 1 s
   "DB_KuKa_MainCtrl.DrillDownload.StepStart" : Bool = PLC DB720_KuKa_MainCtrl.DrillDownload.StepStart AT %DB720.DBX134.4, 1 s
   "DB_KuKa_MainCtrl.DrillUpload.StepStart" : Bool = PLC DB720_KuKa_MainCtrl.DrillUpload.StepStart AT %DB720.DBX144.4, 1 s

HMI tags "Tag_Analog_IN_V4"
   "Analog_In_V4_TP_Cmd" : Word AT %DB1080.DBW0, 1 s
   "Analog_In_V4_Ctrl_Out_Cur_Val_Out" : Real AT %DB1080.DBD0, 1 s
   "Analog_In_V4_Ctrl_IN_TP_PreSetValue" : Real AT %DB1080.DBD0, 1 s
   "Analog_In_V4_Ctrl_IN_TP_AI_Gain" : Real AT %DB1080.DBD0, 1 s
   "Analog_In_V4_Ctrl_IN_TP_AI_OffSet" : Real AT %DB1080.DBD0, 1 s
   "Analog_In_V4_Ctrl_IN_TP_ActualAI_1" : Real AT %DB1080.DBD0, 1 s
   "Analog_In_V4_Ctrl_IN_TP_ActualAI_2" : Real AT %DB1080.DBD0, 1 s
   "Analog_In_V4_Ctrl_IN_TP_ActualAI_Value1" : Real AT %DB1080.DBD0, 1 s
   "Analog_In_V4_Ctrl_IN_TP_ActualAI_Value2" : Real AT %DB1080.DBD0, 1 s

HMI tags "Addr_Analog_IN_V4"
   "DB_AddrRegister_Analog_IN_V4_TP_Cmd" : Int = PLC DB1089_AddrRegister.Analog_IN_V4.TP_Cmd, 1 s
   "DB_AddrRegister_Analog_IN_V4_CTRL_OUT_Cur_Val_Out" : Int = PLC DB1089_AddrRegister.Analog_IN_V4.CTRL_OUT_Cur_Val_Out, 1 s
   "DB_AddrRegister_Analog_IN_V4_CTRL_IN_TP_PreSetValue" : Int = PLC DB1089_AddrRegister.Analog_IN_V4.CTRL_IN_TP_PreSetValue, 1 s
   "DB_AddrRegister_Analog_IN_V4_CTRL_IN_TP_AI_Gain" : Int = PLC DB1089_AddrRegister.Analog_IN_V4.CTRL_IN_TP_AI_Gain, 1 s
   "DB_AddrRegister_Analog_IN_V4_CTRL_IN_TP_AI_OffSet" : Int = PLC DB1089_AddrRegister.Analog_IN_V4.CTRL_IN_TP_AI_OffSet, 1 s
   "DB_AddrRegister_Analog_IN_V4_CTRL_IN_TP_ActualAI_1" : Int = PLC DB1089_AddrRegister.Analog_IN_V4.CTRL_IN_TP_ActualAI_1, 1 s
   "DB_AddrRegister_Analog_IN_V4_CTRL_IN_TP_ActualAI_2" : Int = PLC DB1089_AddrRegister.Analog_IN_V4.CTRL_IN_TP_ActualAI_2, 1 s
   "DB_AddrRegister_Analog_IN_V4_CTRL_IN_TP_ActualAI_Value1" : Int = PLC DB1089_AddrRegister.Analog_IN_V4.CTRL_IN_TP_ActualAI_Value1, 1 s
   "DB_AddrRegister_Analog_IN_V4_CTRL_IN_TP_ActualAI_Value2" : Int = PLC DB1089_AddrRegister.Analog_IN_V4.CTRL_IN_TP_ActualAI_Value2, 1 s
   "DB_AddrRegister_Analog_IN_V4_FBCall_StartAddr" : Int = PLC DB1089_AddrRegister.Analog_IN_V4.FBCall_StartAddr, 1 s
   "DB_AddrRegister_Analog_IN_V4_FBCall_IndexNO" : Int = PLC DB1089_AddrRegister.Analog_IN_V4.FBCall_IndexNO, 1 s

HMI tags "Tag_Analog_Out_V3"
   "Analog_Out_Ctrl_IN_TP_PresetValue" : Real = PLC DB1080_Component.Analog_Out.Ctrl_IN.TP_PresetValue, 1 s
   "Analog_Out_TP_Cmd" : Word = PLC DB1080_Component.Analog_Out.TP_Cmd, 1 s
   "Analog_Out_Ctrl_IN_Target" : Real = PLC DB1080_Component.Analog_Out.Ctrl_IN.Target, 1 s
   "nalog_Out_Ctrl_IN_TP_Offset" : Real = PLC DB1080_Component.Analog_Out.Ctrl_IN.TP_Offset, 1 s
   "Analog_Out_Ctrl_IN_TP_Gain" : Real = PLC DB1080_Component.Analog_Out.Ctrl_IN.TP_Gain, 1 s
   "Analog_Out_Ctrl_IN_TP_ActualAO_1" : Real = PLC DB1080_Component.Analog_Out_1.Ctrl_IN.TP_ActualAI_1, 1 s
   "Analog_Out_Ctrl_IN_TP_ActualAO_2" : Real = PLC DB1080_Component.Analog_Out_1.Ctrl_IN.TP_ActualAI_2, 1 s
   "Analog_Out_Ctrl_IN_TP_ActualAO_Value1" : Real = PLC DB1080_Component.Analog_Out_1.Ctrl_IN.TP_ActualAI_Value1, 1 s
   "Analog_Out_Ctrl_IN_TP_ActualAO_Value2" : Real = PLC DB1080_Component.Analog_Out_1.Ctrl_IN.TP_ActualAI_Value2, 1 s
   "DB_Component.Analog_Out_1.Cmd.Read1" : Bool = PLC DB1080_Component.Analog_Out_1.Cmd.Read1, 1 s
   "DB_Component.Analog_Out_1.Cmd.Read2" : Bool = PLC DB1080_Component.Analog_Out_1.Cmd.Read2, 1 s
   "DB_Component.Analog_Out_1.Confirm" : Bool = PLC DB1080_Component.Analog_Out_1.Confirm, 1 s

discrete alarms
   73: 'ST02.Z01.水平探针缸工作位置故障! / Message__64 / E72', class Alarms, trigger "Err005" bit 8
   4: 'Message__004 / Z06.基本位置故障！Q20.7I21.2 / E3', class Alarms, trigger "Err001" bit 3
   8: 'Message__008 / Z08.基本位置故障！Q21.3I24.5 / E7', class Alarms, trigger "Err001" bit 7
   30: '合格件出料超过2个报警,请确认O圈设备正常! / Z11.基本位置故障！ / E29', class Alarms, trigger "Err002" bit 13
   67: 'Message__067 / Message__74 / E66', class Alarms, trigger "Err005" bit 2
   24: 'Message__068 / Z19.基本位置故障！Q23.1I26.0 / E23', class Alarms, trigger "Err002" bit 7
   27: '合格件出料超过2个报警,请确认O圈设备正常! / Z10.工作位置故障！Q21.6 / E26', class Alarms, trigger "Err002" bit 10
   58: '01.请取下非法工件! / Z34.基本位置故障！Q25.5 / E57', class Alarms, trigger "Err004" bit 9
   62: 'Message__062 / Message__72 / E64', class Alarms, trigger "Err004" bit 13
   87: 'Message__087 / Message__94 / E86', class Alarms, trigger "Err006" bit 6
   143: 'ST04.Z04.水平探针缸工作位置故障! / Message__134 / E142', class Alarms, trigger "Err009" bit 14
   28: '左废料盒已满! / Z10.基本位置故障！Q21.7I26.3 / E27', class Alarms, trigger "Err002" bit 11
   140: 'ST04.Z02.垂直探针缸基本位置故障! / Message__131 / E139', class Alarms, trigger "Err009" bit 11
   42: 'Message__042 / Z22.基本位置故障！Q23.3I22.4 / E41', class Alarms, trigger "Err003" bit 9
   35: 'Message__035 / Z29.工作位置故障！Q24.6I25.1 / E34', class Alarms, trigger "Err003" bit 2
   162: 'Message__162', class Alarms, trigger "Err011" bit 1
   6: 'Message__006 / Z07.基本位置故障！Q21.1I21.0 / E5', class Alarms, trigger "Err001" bit 5
   172: 'Message__172 / Message__163 / E171', class Alarms, trigger "Err011" bit 11
   163: 'Message__163 / Message__170 / E162', class Alarms, trigger "Err011" bit 2
   103: 'Message__103 / Message__110 / E102', class Alarms, trigger "Err007" bit 6
   106: '03.Z01.水平探针缸基本位置故障! / Message__97 / E105', class Alarms, trigger "Err007" bit 9
   115: 'Message__115 / Message__122 / E114', class Alarms, trigger "Err008" bit 2
   7: 'Message__007 / Z08.工作位置故障！Q21.2I24.4 / E6', class Alarms, trigger "Err001" bit 6
   95: 'Message__095 / Message__104 / E96', class Alarms, trigger "Err006" bit 14
   60: '01.工件异常丢失报警！ / Z35.基本位置故障！Q25.7 / E59', class Alarms, trigger "Err004" bit 11
   2: 'Message__002 / Z05.基本位置故障！Q20.5I23.3 / E1', class Alarms, trigger "Err001" bit 1
   179: 'Message__179 / Message__186 / E178', class Alarms, trigger "Err012" bit 2
   57: '01.有疑品件! / Z34.工作位置故障！Q25.4I24.2 / E56', class Alarms, trigger "Err004" bit 8
   94: 'Message__094 / Message__104 / E96', class Alarms, trigger "Err006" bit 13
   9: '设备紧急停止中,请复位！', class Alarms, trigger "Err001" bit 8
   141: 'ST04.Z03.夹紧缸工作位置故障! / Message__132 / E140', class Alarms, trigger "Err009" bit 12
   33: 'Message__033 / Z28.工作位置故障！Q24.2I23.4 / E32', class Alarms, trigger "Err003" bit 0
   148: 'Message__148 / Message__155 / E147', class Alarms, trigger "Err010" bit 3
   114: 'Message__114 / Message__121 / E113', class Alarms, trigger "Err008" bit 1
   37: 'Message__037 / Z32.工作位置故障！Q25.0I25.5 / E36', class Alarms, trigger "Err003" bit 4
   149: 'Message__149 / Message__156 / E148', class Alarms, trigger "Err010" bit 4
   96: 'Message__096 / Message__104 / E96', class Alarms, trigger "Err006" bit 15
   156: 'Message__161', class Alarms, trigger "Err010" bit 11
   25: '转盘夹具ID号错误，请检查编码信号！ / Z09.工作位置故障！Q21.4I24.6 / E24', class Alarms, trigger "Err002" bit 8
   123: 'Message__123 / Message__127 / E119', class Alarms, trigger "Err008" bit 10
   15: 'TCP/IP接收故障报警!', class Alarms, trigger "Err001" bit 14
   61: 'Message__061 / Message__72 / E64', class Alarms, trigger "Err004" bit 12
   66: 'ST02.Z05.下位移笔基本位置故障! / Message__73 / E65', class Alarms, trigger "Err005" bit 1
   171: 'Message__171 / Message__162 / E170', class Alarms, trigger "Err011" bit 10
   38: 'Message__038 / Z32.基本位置故障！Q25.1 / E37', class Alarms, trigger "Err003" bit 5
   136: 'Message__136 / Message__143 / E135', class Alarms, trigger "Err009" bit 7
   155: '04.凹面电压NG! / Message__146 / E154', class Alarms, trigger "Err010" bit 10
   86: 'Message__086 / Message__93 / E85', class Alarms, trigger "Err006" bit 5
   131: 'Message__131 / Message__138 / E130', class Alarms, trigger "Err009" bit 2
   54: 'Message__054 / Message__61 / E53', class Alarms, trigger "Err004" bit 5
   44: 'Message__044 / Z23.基本位置故障！Q23.5I22.0 / E43', class Alarms, trigger "Err003" bit 11
   29: '右废料盒已满！ / Z11.工作位置故障！Q22.0I26.4 / E28', class Alarms, trigger "Err002" bit 12
   64: 'Message__064 / Message__72 / E64', class Alarms, trigger "Err004" bit 15
   181: 'Message__181 / Message__188 / E180', class Alarms, trigger "Err012" bit 4
   99: 'Message__099 / Message__106 / E98', class Alarms, trigger "Err007" bit 2
   18: 'Message__018 / Z16.基本位置故障！Q22.3I20.4 / E17', class Alarms, trigger "Err002" bit 1
   32: 'Message__032 / Z12.基本位置故障！ / E31', class Alarms, trigger "Err002" bit 15
   191: 'Message__191 / Message__182 / E190', class Alarms, trigger "Err012" bit 14
   154: '04.齿面电压NG! / Message__145 / E153', class Alarms, trigger "Err010" bit 9
   75: 'ST02.Z02.垂直探针缸工作位置故障! / Message__66 / E74', class Alarms, trigger "Err005" bit 10
   39: 'Message__039 / Z33.工作位置故障！Q25.2I25.7 / E38', class Alarms, trigger "Err003" bit 6
   128: 'Message__128 / Message__127 / E119', class Alarms, trigger "Err008" bit 15
   184: 'Message__184 / Message__191 / E183', class Alarms, trigger "Err012" bit 7
   22: 'Message__022 / Z18.基本位置故障！Q22.7I20.2 / E21', class Alarms, trigger "Err002" bit 5
   26: '串口读取数据错误! / Z09.基本位置故障！Q21.5 / E25', class Alarms, trigger "Err002" bit 9
   79: 'ST02.Z04.上位移笔工作位置故障! / Message__70 / E78', class Alarms, trigger "Err005" bit 14
   177: 'Message__177 / Message__184 / E176', class Alarms, trigger "Err012" bit 0
   11: '气源未打开，请摁下复位按钮！', class Alarms, trigger "Err001" bit 10
   108: '03.Z02.垂直探针缸基本位置故障! / Message__99 / E107', class Alarms, trigger "Err007" bit 11
   98: 'Message__098 / Message__105 / E97', class Alarms, trigger "Err007" bit 1
   125: 'Message__125 / Message__127 / E119', class Alarms, trigger "Err008" bit 12
   72: 'Message__072 / Message__79 / E71', class Alarms, trigger "Err005" bit 7
   101: 'Message__101 / Message__108 / E100', class Alarms, trigger "Err007" bit 4
   117: 'Message__117 / Message__124 / E116', class Alarms, trigger "Err008" bit 4
   20: 'Message__020 / Z17.基本位置故障！Q22.5I20.0 / E19', class Alarms, trigger "Err002" bit 3
   85: 'Message__085 / Message__92 / E84', class Alarms, trigger "Err006" bit 4
   1: '请先按下开始校验按钮！', class Alarms, trigger "Err001" bit 0
   116: 'Message__116 / Message__123 / E115', class Alarms, trigger "Err008" bit 3
   92: 'Message__092 / Message__104 / E96', class Alarms, trigger "Err006" bit 11
   135: 'Message__135 / Message__142 / E134', class Alarms, trigger "Err009" bit 6
   105: '03.Z01.水平探针缸工作位置故障! / Message__96 / E104', class Alarms, trigger "Err007" bit 8
   120: 'Message__120 / Message__127 / E119', class Alarms, trigger "Err008" bit 7
   97: 'Message__097 / Message__104 / E96', class Alarms, trigger "Err007" bit 0
   152: 'Message__152 / Message__159 / E151', class Alarms, trigger "Err010" bit 5
   84: 'Message__084 / Message__91 / E83', class Alarms, trigger "Err006" bit 3
   91: '02.功能长度测试NG! / Message__82 / E90', class Alarms, trigger "Err006" bit 10
   13: 'PLC与上位机TCP/IP通讯报警!', class Alarms, trigger "Err001" bit 12
   16: '转盘未Ready报警!', class Alarms, trigger "Err001" bit 15
   147: 'Message__147 / Message__154 / E146', class Alarms, trigger "Err010" bit 2
   158: 'Message__161', class Alarms, trigger "Err010" bit 13
   41: 'Message__041 / Z22.工作位置故障！Q23.2 / E40', class Alarms, trigger "Err003" bit 8
   138: 'ST04.Z01.齿面凹面转换缸基本位置故障! / Message__129 / E137', class Alarms, trigger "Err009" bit 9
   93: 'Message__093 / Message__104 / E96', class Alarms, trigger "Err006" bit 12
   110: '03.Z03.升降缸基本位置故障! / Message__120 / E112', class Alarms, trigger "Err007" bit 13
   134: 'Message__134 / Message__141 / E133', class Alarms, trigger "Err009" bit 5
   137: 'ST04.Z01.齿面凹面转换缸工作位置故障! / Message__128 / E136', class Alarms, trigger "Err009" bit 8
   81: 'Message__081 / Message__88 / E80', class Alarms, trigger "Err006" bit 0
   102: 'Message__102 / Message__109 / E101', class Alarms, trigger "Err007" bit 5
   188: 'Message__188 / Message__179 / E187', class Alarms, trigger "Err012" bit 11
   165: 'Message__165 / Message__172 / E164', class Alarms, trigger "Err011" bit 4
   174: 'Message__174 / Message__165 / E173', class Alarms, trigger "Err011" bit 13
   77: 'ST02.Z03.夹紧缸工作位置故障! / Message__68 / E76', class Alarms, trigger "Err005" bit 12
   133: 'Message__133 / Message__140 / E132', class Alarms, trigger "Err009" bit 4
   157: 'Message__161', class Alarms, trigger "Err010" bit 12
   178: 'Message__178 / Message__185 / E177', class Alarms, trigger "Err012" bit 1
   107: '03.Z02.垂直探针缸工作位置故障! / Message__98 / E106', class Alarms, trigger "Err007" bit 10
   88: 'Message__088 / Message__95 / E87', class Alarms, trigger "Err006" bit 7
   70: 'Message__070 / Message__77 / E69', class Alarms, trigger "Err005" bit 5
   17: 'Message__017 / Z16.工作位置故障！Q22.2I20.5 / E16', class Alarms, trigger "Err002" bit 0
   69: 'Message__069 / Message__76 / E68', class Alarms, trigger "Err005" bit 4
   118: 'Message__118 / Message__125 / E117', class Alarms, trigger "Err008" bit 5
   166: 'Message__166 / Message__173 / E165', class Alarms, trigger "Err011" bit 5
   164: 'Message__164 / Message__171 / E163', class Alarms, trigger "Err011" bit 3
   170: 'Message__170 / Message__161 / E169', class Alarms, trigger "Err011" bit 9
   53: 'Message__053 / Message__60 / E52', class Alarms, trigger "Err004" bit 4
   52: 'Message__052 / Message__59 / E51', class Alarms, trigger "Err004" bit 3
   132: 'Message__132 / Message__139 / E131', class Alarms, trigger "Err009" bit 3
   139: 'ST04.Z02.垂直探针缸工作位置故障! / Message__130 / E138', class Alarms, trigger "Err009" bit 10
   189: 'Message__189 / Message__180 / E188', class Alarms, trigger "Err012" bit 12
   12: '气缸操作条件不满足，请检查！', class Alarms, trigger "Err001" bit 11
   176: 'Message__176 / Message__167 / E175', class Alarms, trigger "Err011" bit 15
   68: 'Message__068 / Message__75 / E67', class Alarms, trigger "Err005" bit 3
   90: '02.CR2电阻电容测试NG！ / Message__81 / E89', class Alarms, trigger "Err006" bit 9
   127: 'Message__127 / E119', class Alarms, trigger "Err008" bit 14
   47: 'Message__047 / Z27.工作位置故障！Q24.0I23.1 / E46', class Alarms, trigger "Err003" bit 14
   145: '04.Z05.备用工作位置故障!', class Alarms, trigger "Err010" bit 0
   173: 'Message__173 / Message__164 / E172', class Alarms, trigger "Err011" bit 12
   5: 'Message__005 / Z07.工作位置故障！Q21.0I21.1 / E4', class Alarms, trigger "Err001" bit 4
   50: 'Message__050 / Z27.基本位置故障！Q24.1I23.0 / E47', class Alarms, trigger "Err004" bit 1
   122: 'Message__122 / Message__127 / E119', class Alarms, trigger "Err008" bit 9
   146: '04.Z05.备用基本位置故障!', class Alarms, trigger "Err010" bit 1
   71: 'Message__071 / Message__78 / E70', class Alarms, trigger "Err005" bit 6
   51: 'Message__051 / Message__58 / E50', class Alarms, trigger "Err004" bit 2
   49: 'Message__049 / Z27.基本位置故障！Q24.1I23.0 / E47', class Alarms, trigger "Err004" bit 0
   190: 'Message__190 / Message__181 / E189', class Alarms, trigger "Err012" bit 13
   100: 'Message__100 / Message__107 / E99', class Alarms, trigger "Err007" bit 3
   82: 'Message__082 / Message__89 / E81', class Alarms, trigger "Err006" bit 1
   160: 'Message__161', class Alarms, trigger "Err010" bit 15
   3: 'Message__003 / Z06.工作位置故障！Q20.6I21.3 / E2', class Alarms, trigger "Err001" bit 2
   34: 'Message__034 / Z28.基本位置故障！Q24.3I23.2 / E33', class Alarms, trigger "Err003" bit 1
   130: 'Message__130 / Message__137 / E129', class Alarms, trigger "Err009" bit 1
   183: 'Message__183 / Message__190 / E182', class Alarms, trigger "Err012" bit 6
   169: 'Message__169 / Message__160 / E168', class Alarms, trigger "Err011" bit 8
   43: 'Message__043 / Z23.工作位置故障！Q23.4I22.1 / E42', class Alarms, trigger "Err003" bit 10
   142: 'ST04.Z03.夹紧缸基本位置故障! / Message__133 / E141', class Alarms, trigger "Err009" bit 13
   19: 'Message__019 / Z17.工作位置故障！Q22.4I20.1 / E18', class Alarms, trigger "Err002" bit 2
   31: 'Message__031 / Z12.工作位置故障！Q22.1I26.5 / E30', class Alarms, trigger "Err002" bit 14
   78: 'ST02.Z03.夹紧缸基本位置故障! / Message__69 / E77', class Alarms, trigger "Err005" bit 13
   36: 'Message__036 / Z29.基本位置故障！Q24.7I25.0 / E35', class Alarms, trigger "Err003" bit 3
   111: '03.Z04.夹紧缸工作位置故障! / Message__120 / E112', class Alarms, trigger "Err007" bit 14
   10: '设备气压低，请复位！', class Alarms, trigger "Err001" bit 9
   129: 'Message__129 / Message__136 / E128', class Alarms, trigger "Err009" bit 0
   46: 'Message__046 / Z24.基本位置故障！Q23.7I22.2 / E45', class Alarms, trigger "Err003" bit 13
   65: 'ST02.Z05.下位移笔工作位置故障! / Message__72 / E64', class Alarms, trigger "Err005" bit 0
   144: 'ST04.Z04.水平探针缸基本位置故障! / Message__135 / E143', class Alarms, trigger "Err009" bit 15
   119: 'Message__119 / Message__126 / E118', class Alarms, trigger "Err008" bit 6
   89: '02.CR1电阻电容测试NG！ / Message__80 / E88', class Alarms, trigger "Err006" bit 8
   192: 'Message__192 / Message__183 / E191', class Alarms, trigger "Err012" bit 15
   74: 'ST02.Z01.水平探针缸基本位置故障! / Message__65 / E73', class Alarms, trigger "Err005" bit 9
   56: 'Message__056 / Message__63 / E55', class Alarms, trigger "Err004" bit 7
   151: 'Message__151 / Message__158 / E150', class Alarms, trigger "Err010" bit 6
   113: 'Message__113 / Message__120 / E112', class Alarms, trigger "Err008" bit 0
   185: 'Message__185 / Message__176 / E184', class Alarms, trigger "Err012" bit 8
   63: 'Message__063 / Message__72 / E64', class Alarms, trigger "Err004" bit 14
   161: 'Message__161', class Alarms, trigger "Err011" bit 0
   167: 'Message__167 / Message__174 / E166', class Alarms, trigger "Err011" bit 6
   83: 'Message__083 / Message__90 / E82', class Alarms, trigger "Err006" bit 2
   180: 'Message__180 / Message__187 / E179', class Alarms, trigger "Err012" bit 3
   112: '03.Z04.夹紧缸基本位置故障! / Message__120 / E112', class Alarms, trigger "Err007" bit 15
   23: 'Message__282 / Z19.工作位置故障！Q23.0I26.1 / E22', class Alarms, trigger "Err002" bit 6
   21: 'Message__021 / Z18.工作位置故障！Q22.6I20.3 / E20', class Alarms, trigger "Err002" bit 4
   59: '01.请取下疑品件！ / Z35.工作位置故障！Q25.6I24.1 / E58', class Alarms, trigger "Err004" bit 10
   48: 'Message__048 / Z27.基本位置故障！Q24.1I23.0 / E47', class Alarms, trigger "Err003" bit 15
   104: 'Message__104 / Message__111 / E103', class Alarms, trigger "Err007" bit 7
   126: 'Message__126 / Message__127 / E119', class Alarms, trigger "Err008" bit 13
   121: 'Message__121 / Message__127 / E119', class Alarms, trigger "Err008" bit 8
   175: 'Message__175 / Message__166 / E174', class Alarms, trigger "Err011" bit 14
   187: 'Message__187 / Message__178 / E186', class Alarms, trigger "Err012" bit 10
   76: 'ST02.Z02.垂直探针缸基本位置故障! / Message__67 / E75', class Alarms, trigger "Err005" bit 11
   186: 'Message__186 / Message__177 / E185', class Alarms, trigger "Err012" bit 9
   55: 'Message__055 / Message__62 / E54', class Alarms, trigger "Err004" bit 6
   80: 'ST02.Z04.上位移笔基本位置故障! / Message__71 / E79', class Alarms, trigger "Err005" bit 15
   124: 'Message__124 / Message__127 / E119', class Alarms, trigger "Err008" bit 11
   45: 'Message__045 / Z24.工作位置故障！Q23.6I22.3 / E44', class Alarms, trigger "Err003" bit 12
   159: 'Message__161', class Alarms, trigger "Err010" bit 14
   14: 'TCP/IP发送故障报警!', class Alarms, trigger "Err001" bit 13
   153: 'Message__153 / Message__144 / E152', class Alarms, trigger "Err010" bit 8
   182: 'Message__182 / Message__189 / E181', class Alarms, trigger "Err012" bit 5
   40: 'Message__040 / Z33.基本位置故障！Q25.3 / E39', class Alarms, trigger "Err003" bit 7
   150: 'Message__150 / Message__157 / E149', class Alarms, trigger "Err010" bit 7
   168: 'Message__168 / Message__175 / E167', class Alarms, trigger "Err011" bit 7
   109: '03.Z03.升降缸工作位置故障! / Message__100 / E108', class Alarms, trigger "Err007" bit 12
   193: 'Message__193 / Message__183 / E191', class Alarms, trigger "Err013" bit 0
   194: 'Message__194', class Alarms, trigger "Err013" bit 1
   195: 'Message__195', class Alarms, trigger "Err013" bit 2
   196: 'Message__196', class Alarms, trigger "Err013" bit 3
   197: 'Message__197', class Alarms, trigger "Err013" bit 4
   198: 'Message__198', class Alarms, trigger "Err013" bit 5
   199: 'Message__199', class Alarms, trigger "Err013" bit 6
   200: 'Message__200', class Alarms, trigger "Err013" bit 7
   201: 'ST06.Z05.夹紧缸工作位置故障!', class Alarms, trigger "Err013" bit 8
   202: 'ST06.Z05.夹紧缸基本位置故障!', class Alarms, trigger "Err013" bit 9
   203: 'ST06.Z06.水平探针缸工作位置故障!', class Alarms, trigger "Err013" bit 10
   204: 'ST06.Z06.水平探针缸基本位置故障!', class Alarms, trigger "Err013" bit 11
   205: 'ST06.Z07.垂直探针缸工作位置故障!', class Alarms, trigger "Err013" bit 12
   206: 'ST06.Z07.垂直探针缸基本位置故障!', class Alarms, trigger "Err013" bit 13
   207: 'ST06.Z08.位移笔工作位置故障!', class Alarms, trigger "Err013" bit 14
   208: 'ST06.Z08.位移笔基本位置故障!', class Alarms, trigger "Err013" bit 15
   209: '06.Z05.备用工作位置故障!', class Alarms, trigger "Err014" bit 0
   210: '06.Z05.备用基本位置故障!', class Alarms, trigger "Err014" bit 1
   211: 'Message__211', class Alarms, trigger "Err014" bit 2
   212: 'Message__212', class Alarms, trigger "Err014" bit 3
   213: 'Message__213', class Alarms, trigger "Err014" bit 4
   214: 'Message__214', class Alarms, trigger "Err014" bit 5
   215: 'Message__215', class Alarms, trigger "Err014" bit 6
   216: 'Message__216', class Alarms, trigger "Err014" bit 7
   217: 'Message__216', class Alarms, trigger "Err014" bit 8
   218: 'Message__216', class Alarms, trigger "Err014" bit 9
   219: 'Message__216', class Alarms, trigger "Err014" bit 10
   220: 'Message__216', class Alarms, trigger "Err014" bit 11
   221: 'Message__216', class Alarms, trigger "Err014" bit 12
   222: 'Message__216', class Alarms, trigger "Err014" bit 13
   223: 'Message__216', class Alarms, trigger "Err014" bit 14
   224: 'Message__216', class Alarms, trigger "Err014" bit 15
   225: 'Message__225', class Alarms, trigger "Err015" bit 0
   226: 'Message__226', class Alarms, trigger "Err015" bit 1
   227: 'Message__227', class Alarms, trigger "Err015" bit 2
   228: 'Message__228', class Alarms, trigger "Err015" bit 3
   229: 'Message__229', class Alarms, trigger "Err015" bit 4
   230: 'Message__230', class Alarms, trigger "Err015" bit 5
   231: 'Message__231', class Alarms, trigger "Err015" bit 6
   232: 'Message__232', class Alarms, trigger "Err015" bit 7
   233: 'Message__233', class Alarms, trigger "Err015" bit 8
   234: 'Message__234', class Alarms, trigger "Err015" bit 9
   235: 'Message__235', class Alarms, trigger "Err015" bit 10
   236: 'Message__236', class Alarms, trigger "Err015" bit 11
   237: 'Message__237', class Alarms, trigger "Err015" bit 12
   238: 'Message__238', class Alarms, trigger "Err015" bit 13
   239: 'Message__239', class Alarms, trigger "Err015" bit 14
   240: 'Message__240', class Alarms, trigger "Err015" bit 15
   241: 'Message__241', class Alarms, trigger "Err016" bit 0
   242: 'Message__242', class Alarms, trigger "Err016" bit 1
   243: 'Message__243', class Alarms, trigger "Err016" bit 2
   244: 'Message__244', class Alarms, trigger "Err016" bit 3
   245: 'Message__245', class Alarms, trigger "Err016" bit 4
   246: 'Message__246', class Alarms, trigger "Err016" bit 5
   247: 'Message__247', class Alarms, trigger "Err016" bit 6
   248: 'Message__248', class Alarms, trigger "Err016" bit 7
   249: 'Message__249', class Alarms, trigger "Err016" bit 8
   250: 'Message__250', class Alarms, trigger "Err016" bit 9
   251: 'Message__251', class Alarms, trigger "Err016" bit 10
   252: 'Message__252', class Alarms, trigger "Err016" bit 11
   253: 'Message__253', class Alarms, trigger "Err016" bit 12
   254: 'Message__254', class Alarms, trigger "Err016" bit 13
   255: 'Message__255', class Alarms, trigger "Err016" bit 14
   256: 'Message__256', class Alarms, trigger "Err016" bit 15
   257: 'Message__257', class Alarms, trigger "Err017" bit 0
   258: 'Message__258', class Alarms, trigger "Err017" bit 1
   259: 'Message__259', class Alarms, trigger "Err017" bit 2
   260: 'Message__260', class Alarms, trigger "Err017" bit 3
   261: 'Message__261', class Alarms, trigger "Err017" bit 4
   262: 'Message__262', class Alarms, trigger "Err017" bit 5
   263: 'Message__263', class Alarms, trigger "Err017" bit 6
   264: 'Message__264', class Alarms, trigger "Err017" bit 7
   265: '08.Z01.升降缸工作位置故障!', class Alarms, trigger "Err017" bit 8
   266: '08.Z01.升降缸基本位置故障!', class Alarms, trigger "Err017" bit 9
   267: 'Message__267', class Alarms, trigger "Err017" bit 10
   268: 'Message__268', class Alarms, trigger "Err017" bit 11
   269: 'Message__269', class Alarms, trigger "Err017" bit 12
   270: 'Message__270', class Alarms, trigger "Err017" bit 13
   271: 'Message__271', class Alarms, trigger "Err017" bit 14
   272: 'Message__272', class Alarms, trigger "Err017" bit 15
   273: '08.Z05.备用工作位置故障!', class Alarms, trigger "Err018" bit 0
   274: '08.Z05.备用基本位置故障!', class Alarms, trigger "Err018" bit 1
   275: 'Message__275', class Alarms, trigger "Err018" bit 2
   276: 'Message__276', class Alarms, trigger "Err018" bit 3
   277: 'Message__277', class Alarms, trigger "Err018" bit 4
   278: 'Message__278', class Alarms, trigger "Err018" bit 5
   279: 'Message__279', class Alarms, trigger "Err018" bit 6
   280: 'Message__280', class Alarms, trigger "Err018" bit 7
   281: '下料产品丢失！', class Alarms, trigger "Err018" bit 8
   282: '请清除废料!', class Alarms, trigger "Err018" bit 9
   283: 'Message__281', class Alarms, trigger "Err018" bit 10
   284: '打标数据传输失败！', class Alarms, trigger "Err018" bit 11
   285: '08.Z03.备用工作位置故障!', class Alarms, trigger "Err018" bit 12
   286: '08.Z03.备用基本位置故障!', class Alarms, trigger "Err018" bit 13
   287: '08.Z04.备用工作位置故障!', class Alarms, trigger "Err018" bit 14
   288: '08.Z04.备用基本位置故障!', class Alarms, trigger "Err018" bit 15
   289: 'Message__289', class Alarms, trigger "Err019" bit 0
   290: 'Message__290', class Alarms, trigger "Err019" bit 1
   291: 'Message__291', class Alarms, trigger "Err019" bit 2
   292: 'Message__292', class Alarms, trigger "Err019" bit 3
   293: 'Message__293', class Alarms, trigger "Err019" bit 4
   294: 'Message__294', class Alarms, trigger "Err019" bit 5
   295: 'Message__295', class Alarms, trigger "Err019" bit 6
   296: 'Message__296', class Alarms, trigger "Err019" bit 7
   297: 'ST10.Z01.插销缸工作位置故障!', class Alarms, trigger "Err019" bit 8
   298: 'ST10.Z01.插销缸基本位置故障!', class Alarms, trigger "Err019" bit 9
   299: 'ST10.Z02.测试滑台缸工作位置故障!', class Alarms, trigger "Err019" bit 10
   300: 'ST10.Z02.测试滑台缸基本位置故障!', class Alarms, trigger "Err019" bit 11
   301: 'ST10.Z03.测试升降缸工作位置故障!', class Alarms, trigger "Err019" bit 12
   302: 'ST10.Z03.测试升降缸基本位置故障!', class Alarms, trigger "Err019" bit 13
   303: 'ST10.Z04.滑台推出缸工作位置故障!', class Alarms, trigger "Err019" bit 14
   304: 'ST10.Z04.滑台推出缸基本位置故障!', class Alarms, trigger "Err019" bit 15
   307: '10.工件异常丢失报警！', class Alarms, trigger "Err020" bit 10
   308: '10.气密测试失败!', class Alarms, trigger "Err020" bit 11
   309: '下料产品丢失！', class Alarms, trigger "Err020" bit 8
   310: '请清除废料!', class Alarms, trigger "Err020" bit 9
   311: 'Message__289', class Alarms, trigger "Err020" bit 14
   312: 'Message__289', class Alarms, trigger "Err020" bit 15
   313: 'Message__289', class Alarms, trigger "Err020" bit 12
   314: 'Message__289', class Alarms, trigger "Err020" bit 13
   315: 'Message__291', class Alarms, trigger "Err020" bit 2
   316: 'Message__292', class Alarms, trigger "Err020" bit 3
   317: 'Message__289', class Alarms, trigger "Err020" bit 0
   318: 'Message__290', class Alarms, trigger "Err020" bit 1
   319: 'Message__295', class Alarms, trigger "Err020" bit 6
   320: 'Message__296', class Alarms, trigger "Err020" bit 7
   321: 'Message__293', class Alarms, trigger "Err020" bit 4
   322: 'Message__294', class Alarms, trigger "Err020" bit 5
   323: 'ST11.Z02.下料夹爪缸工作位置故障!', class Alarms, trigger "Err021" bit 10
   324: 'ST11.Z02.下料夹爪缸基本位置故障!', class Alarms, trigger "Err021" bit 11
   325: 'ST11.Z01.下料升降缸工作位置故障!', class Alarms, trigger "Err021" bit 8
   326: 'ST11.Z01.下料升降缸基本位置故障!', class Alarms, trigger "Err021" bit 9
   327: 'Message__289', class Alarms, trigger "Err021" bit 14
   328: 'Message__289', class Alarms, trigger "Err021" bit 15
   329: 'ST11.Z03.废料阻挡缸工作位置故障!', class Alarms, trigger "Err021" bit 12
   330: 'ST11.Z03.废料阻挡缸基本位置故障!', class Alarms, trigger "Err021" bit 13
   331: 'Message__291', class Alarms, trigger "Err021" bit 2
   332: 'Message__292', class Alarms, trigger "Err021" bit 3
   333: 'Message__289', class Alarms, trigger "Err021" bit 0
   334: 'Message__290', class Alarms, trigger "Err021" bit 1
   335: 'Message__295', class Alarms, trigger "Err021" bit 6
   336: 'Message__296', class Alarms, trigger "Err021" bit 7
   337: 'Message__293', class Alarms, trigger "Err021" bit 4
   338: 'Message__294', class Alarms, trigger "Err021" bit 5
   339: 'Message__289', class Alarms, trigger "Err022" bit 10
   340: 'Message__289', class Alarms, trigger "Err022" bit 11
   341: '下料产品丢失！', class Alarms, trigger "Err022" bit 8
   342: '请清除废料!', class Alarms, trigger "Err022" bit 9
   343: 'Message__289', class Alarms, trigger "Err022" bit 14
   344: 'Message__289', class Alarms, trigger "Err022" bit 15
   345: 'Message__289', class Alarms, trigger "Err022" bit 12
   346: 'Message__289', class Alarms, trigger "Err022" bit 13
   347: 'Message__291', class Alarms, trigger "Err022" bit 2
   348: 'Message__292', class Alarms, trigger "Err022" bit 3
   349: 'Message__289', class Alarms, trigger "Err022" bit 0
   350: 'Message__290', class Alarms, trigger "Err022" bit 1
   351: 'Message__295', class Alarms, trigger "Err022" bit 6
   352: 'Message__296', class Alarms, trigger "Err022" bit 7
   353: 'Message__293', class Alarms, trigger "Err022" bit 4
   354: 'Message__294', class Alarms, trigger "Err022" bit 5

text list "Input_地址": 0 'I0.0'; 1 'I0.1'; 2 'I0.2'; 3 'I0.3'; 4 'I0.4'; 5 'I0.5'; 6 'I0.6'; 7 'I0.7'; 10 'I1.0'; 11 'I1.1'; 12 'I1.2'; 13 'I1.3'; 14 'I1.4'; 15 'I1.5'; 16 'I1.6'; 17 'I1.7'; 20 'I2.0'; 21 'I2.1'; 22 'I2.2'; 23 'I2.3'; 24 'I2.4'; 25 'I2.5'; 26 'I2.6'; 27 'I2.7'; 30 'I3.0'; 31 'I3.1'; 32 'I3.2'; 33 'I3.3'; 34 'I3.4'; 35 'I3.5'; 36 'I3.6'; 37 'I3.7'; 40 'I4.0'; 41 'I4.1'; 42 'I4.2'; 43 'I4.3'; 44 'I4.4'; 45 'I4.5'; 46 'I4.6'; 47 'I4.7'; 50 'I5.0'; 51 'I5.1'; 52 'I5.2'; 53 'I5.3'; 54 'I5.4'; 55 'I5.5'; 56 'I5.6'; 57 'I5.7'; 200 'I20.0 / I6.0'; 201 'I20.1 / I6.1'; 202 'I20.2 / I6.2'; 203 'I20.3 / I6.3'; 204 'I20.4 / I6.4'; 205 'I20.5 / I6.5'; 206 'I20.6 / I6.6'; 207 'I20.7 / I6.7'; 210 'I21.0 / I7.0'; 211 'I21.1 / I7.1'; 212 'I21.2 / I20.0'; 213 'I21.3 / I20.1'; 214 'I21.4 / I20.2'; 215 'I21.5 / I20.3'; 216 'I21.6 / I20.4'; 217 'I21.7 / I20.5'; 220 'I22.0'; 221 'I22.1'; 222 'I22.2 / I21.0'; 223 'I22.3 / I21.1'; 224 'I22.4 / I21.2'; 225 'I22.5 / I21.3'; 226 'I22.6 / I21.4'; 227 'I22.7 / I21.5'; 230 'I23.0 / I21.6'; 231 'I23.1'; 232 'I23.2 / I22.0'; 233 'I23.3 / I22.1'; 234 'I23.4 / I22.2'; 235 'I23.5 / I22.3'; 236 'I23.6 / I22.4'; 237 'I23.7'; 240 'I24.0 / I22.6'; 241 'I24.1 / I22.7'; 242 'I24.2 / I23.0'; 243 'I24.3 / I23.1'; 244 'I24.4 / I23.2'; 245 'I24.5 / I23.3'; 246 'I24.6 / I23.4'; 247 'I24.7 / I23.5'; 250 'I25.0 / I23.6'; 251 'I25.1 / I23.7'; 252 'I25.2 / I24.0'; 253 'I25.3 / I24.1'; 254 'I25.4 / I24.2'; 255 'I25.5 / I24.3'; 256 'I25.6 / I24.4'; 257 'I25.7 / I24.5'; 260 'I26.0 / I24.6'; 261 'I26.1 / I24.7'; 262 'I26.2 / I25.0'; 263 'I26.3 / I25.1'; 264 'I26.4 / I25.2'; 265 'I26.5 / I25.3'; 266 'I26.6 / I25.4'; 267 'I26.7 / I25.5'; 270 'I27.0 / I25.6'; 271 'I27.1 / I25.7'; 272 'I27.2 / I26.0'; 273 'I27.3 / I26.1'; 274 'I27.4 / I26.2'; 275 'I27.5 / I26.3'; 276 'I27.6 / I26.4'; 277 'I27.7 / I26.5'; 280 'I28.0 / I26.6'; 281 'I28.1'; 282 'I28.2'; 283 'I28.3'; 284 'I28.4'; 285 'I28.5'; 286 'I28.6'; 287 'I28.7'; 290 'I29.0'; 291 'I29.1'; 292 'I29.2'; 293 'I29.3'; 294 'I29.4'; 295 'I29.5'; 296 'I29.6'; 297 'I29.7'; 300 'I30.0'; 301 'I30.1'; 302 'I30.2'; 303 'I30.3'; 304 'I30.4'; 305 'I30.5'; 306 'I30.6'; 307 'I30.7'; 310 'I31.0'; 311 'I31.1'; 312 'I31.2'; 313 'I31.3'; 314 'I31.4'; 315 'I31.5'; 316 'I31.6'; 317 'I31.7'; 60 'I6.0'; 61 'I6.1'; 62 'I6.2'; 63 'I6.3'; 64 'I6.4'; 65 'I6.5'; 66 'I6.6'; 67 'I6.7'; 71 'I7.1'; 70 'I7.0'; 77 'I7.7'; 76 'I7.6'; 75 'I7.5'; 74 'I7.4'; 73 'I7.3'; 72 'I7.2'; 320 'I32.0'; 321 'I32.1'; 322 'I32.2'; 323 'I32.3'; 324 'I32.4'; 325 'I32.5'; 326 'I32.6'; 327 'I32.7'; 330 'I33.0'; 331 'I33.1'; 332 'I33.2'; 333 'I33.3'; 334 'I33.4'; 335 'I33.5'; 336 'I33.6'; 337 'I33.7'; 340 'I34.0'; 341 'I34.1'; 342 'I34.2'; 343 'I34.3'; 344 'I34.4'; 345 'I34.5'; 346 'I34.6'; 347 'I34.7'; 350 'I35.0'; 351 'I35.1'; 352 'I35.2'; 353 'I35.3'; 354 'I35.4'; 355 'I35.5'; 356 'I35.6'; 357 'I35.7'

text list "Cylinder_Name": 1 '推力气缸 原点位Z01'; 2 '辅助气缸 原点位Z02'; 3 '左防尘盖夹紧缸 原点位Z03'; 4 '右防尘盖夹紧缸 原点位Z04'; 5 '枪钻上电关 开Z05'; 6 '水泥板吹气 关闭Z06'; 7 '快换盘锁紧 锁紧Z07'; 8 '参数 原点位Z08'; 9 '清零 读取Z09'; 10 '18V 原点位Z10'; 11 '24V 原点位Z11'; 12 '36V 原点位Z12'; 13 '03.备用 原点位Z03'; 14 '03.备用 原点位Z04'; 15 '03.备用 原点位Z05'

text list "按钮1": 0 '\\ 公共 操作'; 200..299 '主 画面'; 300..399 '\\ 仪器 程序'; 400..499 '\\ / /'

text list "Cylinder_QExt": 1 'Q20.0'; 2 'Q20.3'; 3 'Q20.2'; 4 ''; 5 'Q20.5'; 6 'Q20.7'; 7 'Q23.0'; 8 ''; 9 ''; 10 ''; 11 ''; 12 ''; 13 ''; 14 ''; 15 ''; 16 'Q21.2'; 17 'Q23.2'; 18 ''; 19 ''; 20 ''; 21 'Q22.2'; 22 'Q22.4'; 23 'Q22.6'; 24 'Q23.4'; 25 ''; 26 'Q20.2'; 27 ''; 28 ''; 29 ''; 30 ''; 31 'Q23.6'; 32 'Q24.0'; 33 'Q24.2'; 34 'Q24.4'; 35 'Q24.6'; 36 'Q25.0'; 37 'Q25.2'; 38 'Q25.4'; 39 ''; 40 ''; 41 ''; 42 ''; 43 ''

text list "Cylinder_QRet": 1 'Q20.1'; 2 ''; 3 ''; 4 ''; 5 'Q20.4'; 6 'Q20.6'; 7 'Q23.1'; 8 ''; 9 ''; 10 ''; 11 ''; 12 ''; 13 ''; 14 ''; 15 ''; 16 'Q21.3'; 17 'Q23.3'; 18 ''; 19 ''; 20 ''; 21 'Q22.3'; 22 'Q22.5'; 23 'Q22.7'; 24 'Q23.5'; 25 ''; 26 'Q20.3'; 27 ''; 28 ''; 29 ''; 30 ''; 31 'Q23.7'; 32 'Q24.1'; 33 'Q24.3'; 34 'Q24.5'; 35 'Q24.7'; 36 'Q25.1'; 37 'Q25.3'; 38 'Q25.5'; 39 ''; 40 ''; 41 ''; 42 ''; 43 ''

text list "气缸运行条件": 0 '条件如下：'; 0 '欢迎使用本系统！ / P10000'; 1 '条件如下： 1: OverAllPmt=ON'; 2 '条件如下：'; 3 '条件如下： 1: OverAllPmt=ON'; 4 '条件如下：'; 5 '条件如下： 1: OverAllPmt=ON'; 6 '条件如下：'; 7 '条件如下： 1: OverAllPmt=ON'; 8 '条件如下：'; 9 '条件如下： 1: OverAllPmt=ON'; 10 '条件如下：'; 11 '条件如下： 1: OverAllPmt=ON'; 12 ''; 13 ''; 14 ''; 15 ''; 16 ''; 17 ''; 18 ''; 19 ''; 20 ''; 21 ''; 22 ''; 23 ''; 24 ''; 25 ''; 26 ''; 27 ''; 28 ''; 29 ''; 30 ''; 31 ''; 32 ''; 33 ''; 34 ''; 35 ''; 36 ''; 37 ''; 38 '条件如下：'; 39 '条件如下： 1: OverAllPmt=ON 2: Z21.RetPos=ON 3: Z22.RetPos=ON 4: Z23.ExtPos=ON'; 40 '条件如下： 1: OverAllPmt=ON'; 41 '条件如下： 1: OverAllPmt=ON 2: (Z20.ExtPos=ON或者Z20.RetPos=ON) 3: Z23.ExtPos=ON'; 42 '条件如下： 1: OverAllPmt=ON'; 43 '条件如下： 1: OverAllPmt=ON 2: (Z20.ExtPos=ON或者Z20.RetPos=ON) 3: Z23.ExtPos=ON'; 44 '条件如下： 1: OverAllPmt=ON 2: Z21.RetPos=ON 3: Z22.RetPos=ON'; 45 '条件如下： 1: OverAllPmt=ON'; 46 '条件如下：'; 47 '条件如下： 1: OverAllPmt=ON'; 48 '条件如下：'; 49 '条件如下： 1: OverAllPmt=ON'; 50 '条件如下：'; 51 '条件如下： 1: OverAllPmt=ON'; 52 ''; 53 ''; 54 ''; 55 ''; 56 ''; 57 ''; 58 '条件如下：'; 59 '条件如下： 1: OverAllPmt=ON'

text list "按钮5": 0 '/ /'; 200..299 '备用'; 300..399 '备用 系统 设定'; 400..499 '备用'

text list "Cylinder_IRet": 1 'I20.0 / I25.3'; 2 'I24.7'; 3 'I21.6'; 4 ''; 5 'I23.4'; 6 'I21.3'; 7 'I24.0'; 8 ''; 9 ''; 10 ''; 11 ''; 12 ''; 13 ''; 14 ''; 15 ''; 16 'I20.5'; 17 'I25.0'; 18 ''; 19 ''; 20 ''; 21 'I26.0'; 22 'I26.2'; 23 'I26.4'; 24 'I25.2'; 25 ''; 26 'I20.3'; 27 ''; 28 ''; 29 ''; 30 ''; 31 'I29.0'; 32 'I29.2'; 33 'I29.4'; 34 'I29.7'; 35 'I30.0'; 36 'I30.3'; 37 'I30.4'; 38 'I30.7'; 39 ''; 40 ''

text list "Cylinder_IExt": 1 'I20.1 / I25.3'; 2 'I24.7'; 3 'I21.6'; 4 ''; 5 ''; 6 'I21.3'; 7 'I24.1'; 8 ''; 9 ''; 10 ''; 11 ''; 12 ''; 13 ''; 14 ''; 15 ''; 16 'I20.4'; 17 'I25.1'; 18 ''; 19 'I25.3'; 20 ''; 21 'I26.1'; 22 'I26.3'; 23 ''; 24 'I25.3'; 25 ''; 26 ''; 27 ''; 28 ''; 29 ''; 30 ''; 31 'I29.1'; 32 'I29.3'; 33 'I29.5'; 34 'I29.6'; 35 'I30.1'; 36 'I30.2'; 37 'I30.5'; 38 'I30.6'; 39 ''; 40 ''; 41 ''; 42 ''; 43 ''

text list "操作提示": 0 '气缸操作被禁止，请检查安全条件！'; 1 '设备处于单步模式，请注意安全！'; 2 '设备已经开始清空，请等待！'; 3 '等待循环结束，暂停自动模式中！'; 4 '开始安全门旁路,等待各流程结束!'; 5 '请启动设备！'; 6 '模式来自触摸屏，调试中！'; 7 '光幕被遮,注意安全!'; 8 '请摁下自动模式启动按钮！'; 9 '请求上位机参数录入...'; 10 '请开始换夹具...'; 11 '请求上位机参数录入...'; 12 '换爪运行中'; 13 '水平方向钻入运行中'; 14 '向上方向钻入运行中'; 15 '向下方向钻入运行中'; 16 '检查钻头运行中'; 17 '清洁运行中'; 18 '换爪位置'; 19 '水平方向钻入位置'; 20 '向上方向钻入位置'; 21 '向下方向钻入位置'; 22 '检查钻头位置'; 23 '请求钻孔'; 24 '请求停止钻孔'; 25 '清洁位置'; 26 '换爪完成'; 27 '水平方向钻入完成'; 28 '向上方向钻入完成'; 29 '向下方向钻入完成'; 30 '检查钻头完成'; 31 ''; 32 '01.Z01.解锁缸到工作位置...'; 33 '01.Z01.解锁缸到基本位置...'; 34 '01.Z02.备用到工作位置...'; 35 '01.Z02.备用到基本位置...'; 36 '01.Z03.备用到工作位置...'; 37 '01.Z03.备用到基本位置...'; 38 '01.Z04.备用到工作位置...'; 39 '01.Z04.备用到基本位置...'; 40 '01.Z05.备用到工作位置...'; 41 '01.Z05.备用到基本位置...'; 42 ''; 43 ''; 44 ''; 45 ''; 46 ''; 47 ''; 48 ''; 49 ''; 50 ''; 51 ''; 52 '等待推力缸完全释放'; 53 '等待推力缸完全释放'; 54 '等待推力缸完全释放'; 55 ''; 56 ''; 57 ''; 58 ''; 59 ''; 60 ''; 61 ''; 62 ''; 63 ''; 64 'ST02.Z01.水平探针缸到工作位置...'; 65 'ST02.Z01.水平探针缸到基本位置...'; 66 'ST02.Z02.垂直探针缸到工作位置...'; 67 'ST02.Z02.垂直探针缸到基本位置...'; 68 'ST02.Z03.夹紧缸到工作位置...'; 69 'ST02.Z03.夹紧缸到基本位置...'; 70 'ST02.Z04.上位移笔到工作位置...'; 71 'ST02.Z04.上位移笔到基本位置...'; 72 'ST02.Z05.下位移笔到工作位置...'; 73 'ST02.Z05.下位移笔到基本位置...'; 74 ''; 75 ''; 76 ''; 77 ''; 78 ''; 79 ''; 80 '02.等待上位机电阻电容反馈结果清零...'; 81 '02.等待上位机功能长度反馈结果清零...'; 82 '02.等待串口通讯空闲...'; 83 '02.等待串口读取数据开始...'; 84 '02.等待串口读取数据结束...'; 85 '02.CR1测试中...'; 86 '02.CR2测试中...'; 87 '02.功能长度测试中...'; 88 ''; 89 ''; 90 ''; 91 ''; 92 ''; 93 ''; 94 ''; 95 ''; 96 '03.Z01.水平探针缸到工作位置...'; 97 '03.Z01.水平探针缸到基本位置...'; 98 '03.Z02.垂直探针缸到工作位置...'; 99 '03.Z02.垂直探针缸到基本位置...'; 100 '03.Z03.升降缸到工作位置...'; 101 '03.Z03.升降缸到基本位置...'; 102 '03.Z04.夹紧缸到工作位置...'; 103 '03.Z04.夹紧缸到基本位置...'; 104 '03.Z05.备用到工作位置...'; 105 '03.Z05.备用到基本位置...'; 106 ''; 107 ''; 108 ''; 109 ''; 110 ''; 111 ''; 112 ''; 113 ''; 114 ''; 115 ''; 116 ''; 117 ''; 118 ''; 119 ''; 120 ''; 121 ''; 122 ''; 123 ''; 124 ''; 125 ''; 126 ''; 127 ''; 128 'ST04.Z01.齿面凹面转换缸到工作位置...'; 129 'ST04.Z01.齿面凹面转换缸到基本位置...'; 130 'ST04.Z02.垂直探针缸到工作位置...'; 131 'ST04.Z02.垂直探针缸到基本位置...'; 132 'ST04.Z03.夹紧缸到工作位置...'; 133 'ST04.Z03.夹紧缸到基本位置...'; 134 'ST04.Z04.水平探针缸到工作位置...'; 135 'ST04.Z04.水平探针缸到基本位置...'; 136 '04.Z05.水平探针缸到工作位置...'; 137 '04.Z05.水平探针缸到基本位置...'; 138 ''; 139 ''; 140 ''; 141 ''; 142 ''; 143 ''; 144 ''; 145 ''; 146 ''; 147 ''; 148 ''; 149 ''; 150 ''; 151 ''; 152 ''; 153 ''; 154 ''; 155 ''; 156 ''; 157 ''; 158 ''; 159 ''; 160 '05.Z01.备用到工作位置...'; 161 '05.Z01.备用到基本位置...'; 162 '05.Z02.备用到工作位置...'; 163 '05.Z02.备用到基本位置...'; 164 '05.Z03.备用到工作位置...'; 165 '05.Z03.备用到基本位置...'; 166 '05.Z04.备用到工作位置...'; 167 '05.Z04.备用到基本位置...'; 168 '05.Z05.备用到工作位置...'; 169 '05.Z05.备用到基本位置...'; 170 ''; 171 ''; 172 ''; 173 ''; 174 ''; 175 ''; 176 '05.等待上位机反馈结果清零...'; 177 '05.等待串口通讯空闲...'; 178 '05.等待串口读取数据开始...'; 179 '05.等待串口读取数据结束...'; 180 ''; 181 ''; 182 ''; 183 ''; 184 ''; 185 ''; 186 ''; 187 ''; 188 ''; 189 ''; 190 ''; 191 ''; 192 'ST06.Z01.夹紧缸工作位置故障!'; 193 'ST06.Z01.夹紧缸基本位置故障!'; 194 'ST06.Z02.水平探针缸工作位置故障!'; 195 'ST06.Z02.水平探针缸基本位置故障!'; 196 'ST06.Z03.垂直探针缸工作位置故障!'; 197 'ST06.Z03.垂直探针缸基本位置故障!'; 198 'ST06.Z04.位移笔工作位置故障!'; 199 'ST06.Z04.位移笔基本位置故障!'; 200 '06.Z05.备用到工作位置...'; 201 '06.Z05.备用到基本位置...'; 202 ''; 203 ''; 204 ''; 205 ''; 206 ''; 207 '06.工件OK/NG结果请求中...'; 208 '06.等待打标机空闲,写入打标内容...'; 209 '06.写入打标变量内容...'; 210 '06.等待打标机空闲,启动打标...'; 211 '06.启动打标...'; 212 '06.等待上位机反馈结果清零...'; 213 ''; 214 ''; 215 ''; 216 ''; 217 ''; 218 ''; 219 ''; 220 ''; 221 ''; 222 ''; 223 ''; 224 '07.Z01.插销缸到工作位置...'; 225 '07.Z01.插销缸到基本位置...'; 226 '07.Z02.压紧缸到工作位置...'; 227 '07.Z02.压紧缸到基本位置...'; 228 '07.Z03.测试缸到工作位置...'; 229 '07.Z03.测试缸到基本位置...'; 230 '07.Z04.滑台推出缸到工作位置...'; 231 '07.Z04.滑台推出缸到基本位置...'; 232 '07.Z05.下料滑台缸到工作位置...'; 233 '07.Z05.下料滑台缸到基本位置...'; 250 ''; 251 ''; 252 ''; 253 ''; 254 ''; 255 ''; 256 '08.Z01.升降缸到工作位置...'; 257 '08.Z01.升降缸到基本位置...'; 258 ''; 259 ''; 260 ''; 261 ''; 262 ''; 263 ''; 264 ''; 265 ''; 266 ''; 267 ''; 268 ''; 269 ''; 270 ''; 271 ''; 272 ''; 273 ''; 274 ''; 275 ''; 276 ''; 277 ''; 278 ''; 279 ''; 280 ''; 281 ''; 282 ''; 283 ''; 284 ''; 285 ''; 286 ''; 287 ''; 288 'ST10.Z01.插销缸到工作位置...'; 289 'ST10.Z01.插销缸到基本位置...'; 290 'ST10.Z02.测试滑台缸到工作位置...'; 291 'ST10.Z02.测试滑台缸到基本位置...'; 292 'ST10.Z03.测试升降缸到工作位置...'; 293 'ST10.Z03.测试升降缸到基本位置...'; 294 'ST10.Z04.滑台推出缸到工作位置...'; 295 'ST10.Z04.滑台推出缸到基本位置...'; 296 'ST10.Z05.下料滑台缸到工作位置...'; 297 'ST10.Z05.下料滑台缸到基本位置...'; 298 ''; 299 ''; 300 ''; 301 ''; 302 ''; 1000 '设备不在原点,需要复位!'; 1001 '请摁下自动模式启动按钮！'; 1002 '安全门旁路，注意安全！'; 1003 '安全门电磁线圈锁定失败！'; 1004 '上位机通讯失败！'; 1005 ''; 1006 ''; 1007 ''; 1008 ''; 1009 ''; 1010 ''; 1011 ''; 1012 ''; 1013 ''; 1014 ''; 1015 ''; 1016 ''; 1017 ''; 1018 ''; 1019 ''; 1020 ''; 1021 ''; 1022 ''; 1023 ''; 1024 ''; 1025 ''; 1026 ''; 1027 ''; 1028 ''; 1029 ''; 1030 ''; 1031 ''; 1032 ''; 1033 ''; 1034 ''; 1035 ''; 1036 ''; 1037 ''; 1038 ''; 1039 ''; 1040 ''; 1041 ''; 1042 ''; 1043 ''; 1044 ''; 1045 ''; 1046 ''; 1047 ''; 1048 '请取下合格件!'; 1049 '请取下疑品件!'; 1050 ''; 1051 ''; 1052 ''; 1053 ''; 1054 ''; 1055 ''; 1056 ''; 1057 ''; 1058 ''; 1059 ''; 1060 ''; 1061 ''; 1062 ''; 1063 ''; 1064 ''; 1065 ''; 1066 ''; 1067 ''; 1068 ''; 1069 ''; 1070 ''; 1071 ''; 1072 ''; 1073 ''; 1074 ''; 1075 ''; 1076 ''; 1077 ''; 1078 ''; 1079 ''; 1080 ''; 1081 ''; 1082 ''; 1083 ''; 1084 ''; 1085 ''; 1086 ''; 1087 ''; 1088 ''; 1089 ''; 1090 ''; 1091 ''; 1092 ''; 1093 ''; 1094 ''; 1095 ''; 1096 ''; 1097 ''; 1098 ''; 1099 ''; 1100 ''; 1101 ''; 1102 ''; 1103 ''; 1104 ''; 1105 ''; 1106 ''; 1107 ''; 1108 ''; 1109 ''; 1110 ''; 1111 ''; 1112 ''; 1113 ''; 1114 ''; 1115 ''; 1116 ''; 1117 ''; 1118 ''; 1119 ''; 1120 ''; 1121 ''; 1122 ''; 1123 ''; 1124 ''; 1125 ''; 1126 ''; 1127 ''; 1128 ''; 1129 ''; 1130 ''; 1131 ''; 1132 ''; 1133 ''; 1134 ''; 1135 ''; 1136 ''; 1137 ''; 1138 ''; 1139 ''; 1140 ''; 1141 ''; 1142 ''; 1143 ''; 1144 ''; 1145 ''; 1146 ''; 1147 ''; 1148 ''; 1149 ''; 1150 ''; 1151 ''; 1152 ''; 1153 ''; 1154 ''; 1155 ''; 1156 ''; 1157 ''; 1158 ''; 1159 ''; 1160 ''; 1161 ''; 1162 ''; 1163 ''; 1164 ''; 1165 ''; 1166 ''; 1167 ''; 1168 ''; 1169 ''; 1170 ''; 1171 ''; 1172 ''; 1173 ''; 1174 ''; 1175 ''; 1176 ''; 1177 ''; 1178 ''; 1179 ''; 1180 ''; 1181 ''; 1182 ''; 1183 ''; 1184 ''; 1185 ''; 1186 ''; 1187 ''; 1188 ''; 1189 ''; 1190 ''; 1191 ''; 1192 ''; 1193 ''; 1194 ''; 1195 ''; 1196 ''; 1197 ''; 1198 ''; 1199 ''; 1200 ''; 1201 ''; 1202 ''; 1203 ''; 1204 ''; 1205 ''; 1206 ''; 1207 ''; 1208 ''; 1209 ''; 1210 ''; 1211 ''; 1212 ''; 1213 ''; 1214 ''; 1215 ''; 1216 ''; 1217 ''; 1218 ''; 1219 ''; 1220 ''; 1221 ''; 1222 ''; 1223 ''; 1224 ''; 1225 ''; 1226 ''; 1227 ''; 1228 ''; 1229 ''; 1230 ''; 1231 ''; 1232 ''; 1233 ''; 1234 ''; 1235 ''; 1236 ''; 1237 ''; 1238 ''; 1239 ''; 1240 ''; 1241 ''; 1242 ''; 1243 ''; 1244 ''; 1245 ''; 1246 ''; 1247 ''; 1248 ''; 1249 ''; 1250 ''; 1251 ''; 1252 ''; 1253 ''; 1254 ''; 1255 ''; 1256 ''; 1257 ''; 1258 ''; 1259 ''; 1260 ''; 1261 ''; 1262 ''; 1263 ''; 1264 ''; 1265 ''; 1266 ''; 1267 ''; 1268 ''; 1269 ''; 1270 ''; 1271 ''; 1272 ''; 1273 ''; 1274 ''; 1275 ''; 1276 ''; 1277 ''; 1278 ''; 1279 ''; 1280 ''; 1281 ''; 1282 ''; 1283 ''; 1284 ''; 1285 ''; 1286 ''; 1287 ''; 1288 ''; 1289 ''; 1290 ''; 1291 ''; 1292 ''; 1293 ''; 1294 ''; 1295 ''; 1296 ''; 1297 ''; 1298 ''; 1299 ''; 1300 ''; 1301 ''; 1302 ''; 2000 '设备紧急停止中,请复位！'; 2001 '设备气压低，请复位！'; 2002 '气源未打开，请摁下复位按钮！'; 2003 '气缸操作条件不满足，请检查！'; 2004 '上位机急停！'; 2005 '打孔超时！'; 2006 '推力缸初始位置不正确！'; 2007 ''; 2008 ''; 2009 '机器人未准备好！'; 2010 '操作盒急停NOK'; 2011 '机器人急停按钮NOK'; 2012 '温控器报警'; 2013 '围栏内侧急停NOK'; 2014 '水泥块击打框架急停NOK'; 2015 'Beeper_17'; 2016 '电源夹具ID号错误，请检查夹具！'; 2017 ''; 2018 ''; 2019 ''; 2020 ''; 2021 ''; 2022 '光幕被遮，确认安全后复位！'; 2023 '信号夹具ID号错误，请检查夹具！'; 2024 '水平水泥板已打完，请更换水泥板！'; 2025 '垂直向上水泥板已打完，请更换水泥板！'; 2026 '垂直向下水泥板已打完，请更换水泥板！'; 2027 '批头长度错误，请更换！'; 2028 ''; 2029 ''; 2030 ''; 2031 ''; 2032 'Z01.推力气缸工作位置故障!'; 2033 'Z01.推力气缸基本位置故障!'; 2034 'Z02.辅助气缸工作位置故障!'; 2035 'Z02.辅助气缸基本位置故障!'; 2036 'Z03.左防尘盖夹紧缸工作位置故障!'; 2037 'Z03.左防尘盖夹紧缸基本位置故障!'; 2038 'Z04.右防尘盖夹紧缸工作位置故障!'; 2039 'Z04.右防尘盖夹紧缸基本位置故障!'; 2040 'Z05.枪电源工作位置故障!'; 2041 'Z05.枪电源基本位置故障!'; 2042 'Z06.水泥板吹气工作位置故障!'; 2043 'Z06.水泥板吹气基本位置故障!'; 2044 'Z07.快换盘锁紧工作位置故障!'; 2045 'Z07.快换盘锁紧基本位置故障!'; 2046 ''; 2047 ''; 2048 ''; 2049 ''; 2050 ''; 2051 ''; 2052 ''; 2053 ''; 2054 ''; 2055 ''; 2056 ''; 2057 ''; 2058 ''; 2059 ''; 2060 ''; 2061 ''; 2062 ''; 2063 ''; 2349 '欢迎使用本系统！'; 310 ''; 309 ''; 308 ''; 307 ''; 305 ''; 306 ''; 304 ''; 303 ''; 348 ''; 327 ''; 326 ''; 311 ''; 325 'ST11.Z03.废料阻挡缸到基本位置...'; 312 ''; 324 'ST11.Z03.废料阻挡缸到工作位置...'; 323 'ST11.Z02.下料夹爪缸到基本位置...'; 322 'ST11.Z02.下料夹爪缸到工作位置...'; 321 'ST11.Z01.下料升降缸到基本位置...'; 320 'ST11.Z01.下料升降缸到工作位置...'; 313 ''; 319 ''; 318 ''; 317 ''; 316 ''; 315 ''; 314 ''; 347 ''; 346 ''; 345 ''; 344 ''; 343 ''; 342 ''; 328 ''; 341 ''; 340 ''; 339 ''; 338 ''; 337 ''; 336 ''; 335 ''; 330 ''; 329 ''; 334 ''; 333 ''; 332 ''; 331 ''; 248 ''; 247 ''; 246 ''; 235 ''; 234 ''; 245 ''; 244 ''; 243 ''; 242 ''; 241 ''; 240 ''; 238 ''; 239 ''; 237 ''; 236 ''; 249 ''

text list "按钮4": 0 '\\ / /'; 200..299 'IO Check'; 300..399 '\\ / 备用'; 400..499 '\\ / 备用'

text list "按钮2": 0 '\\ 机器 人'; 200..299 '\\ 统计 信息'; 300..399 '\\ 伺服 位置'; 400..499 '\\ / /'

text list "气缸条件页名": 1 '01.旋转缸 ( Z01 ) 工作位置条件'; 2 '01.旋转缸 ( Z01 ) 原点位置条件'; 3 '01.真空 ( Z02 ) 工作位置条件'; 4 '01.真空 ( Z02 ) 原点位置条件'; 5 '02.真空 ( Z03 ) 工作位置条件'; 6 '02.真空 ( Z03 ) 原点位置条件'; 7 ''; 8 ''; 9 '02.升降缸 ( Z05 ) 工作位置条件'; 10 '02.升降缸 ( Z05 ) 原点位置条件'; 11 '02.伸出1缸 ( Z06 ) 工作位置条件'; 12 '02.伸出1缸 ( Z06 ) 原点位置条件'; 13 '02.伸出2缸 ( Z07 ) 工作位置条件'; 14 '02.伸出2缸 ( Z07 ) 原点位置条件'; 15 '02.送料长缸 ( Z08 ) 工作位置条件'; 16 '02.送料长缸 ( Z08 ) 原点位置条件'; 17 '02.送料短缸 ( Z09 ) 工作位置条件'; 18 '02.送料短缸 ( Z09 ) 原点位置条件'; 19 '02.送料升降缸 ( Z10 ) 工作位置条件'; 20 '02.送料升降缸 ( Z10 ) 原点位置条件'; 21 '02.送料夹爪缸 ( Z11 ) 工作位置条件'; 22 '02.送料夹爪缸 ( Z11 ) 原点位置条件'; 23 '02.剥料缸 ( Z12 ) 工作位置条件'; 24 '02.剥料缸 ( Z12 ) 原点位置条件'; 25 '振动料斗 ( Z13 ) 工作位置条件'; 26 '振动料斗 ( Z13 ) 原点位置条件'; 27 ''; 28 ''; 29 ''; 30 ''; 31 '03.压紧缸 ( Z16 ) 工作位置条件'; 32 '03.压紧缸 ( Z16 ) 原点位置条件'; 33 '03.伸出1缸 ( Z17 ) 工作位置条件'; 34 '03.伸出1缸 ( Z17 ) 原点位置条件'; 35 '03.伸出2缸 ( Z18 ) 工作位置条件'; 36 '03.伸出2缸 ( Z18 ) 原点位置条件'; 37 '03.测试缸 ( Z19 ) 工作位置条件'; 38 '03.测试缸 ( Z19 ) 原点位置条件'; 39 ''; 40 ''; 41 ''; 42 ''; 43 '05.压紧缸 ( Z22 ) 工作位置条件'; 44 '05.压紧缸 ( Z22 ) 原点位置条件'; 45 '05.伸出1缸 ( Z23 ) 工作位置条件'; 46 '05.伸出1缸 ( Z23 ) 原点位置条件'; 47 '05.伸出2缸 ( Z24 ) 工作位置条件'; 48 '05.伸出2缸 ( Z24 ) 原点位置条件'; 49 ''; 50 ''; 51 ''; 52 ''; 53 '06.压紧缸 ( Z27 ) 工作位置条件'; 54 '06.压紧缸 ( Z27 ) 原点位置条件'; 55 '06.热烫缸 ( Z28 ) 工作位置条件'; 56 '06.热烫缸 ( Z28 ) 原点位置条件'; 57 '06.检测缸 ( Z29 ) 工作位置条件'; 58 '06.检测缸 ( Z29 ) 原点位置条件'; 59 ''; 60 ''; 61 ''; 62 ''; 63 '上料皮带挡料1缸 ( Z32 ) 工作位置条件'; 64 '上料皮带挡料1缸 ( Z32 ) 原点位置条件'; 65 '上料皮带挡料2缸 ( Z33 ) 工作位置条件'; 66 '上料皮带挡料2缸 ( Z33 ) 原点位置条件'; 67 '下料皮带挡料1缸 ( Z34 ) 工作位置条件'; 68 '下料皮带挡料1缸 ( Z34 ) 原点位置条件'; 69 '下料皮带挡料2缸 ( Z35 ) 工作位置条件'; 70 '下料皮带挡料2缸 ( Z35 ) 原点位置条件'; 71 '离子吹气 ( Z36 ) 工作位置条件'; 72 '离子吹气 ( Z36 ) 原点位置条件'

text list "按钮3": 0 '\\ 伺服 操作'; 200..299 '\\ 校验 信息'; 300..399 '\\ 仪器 程序'; 400..499 '\\ / 备用'

text list "工作模式": 0 '手动模式'; 1 '校验模式 / 自动模式'; 2 '单步模式'; 3 '自动模式 / 校验模式'; 4 '系统紧停'; 5 '气压低 / 调试模式'

text list "功能选择": 0 '开启'; 1 '关闭'

text list "启用禁用": 0 '启用'; 1 '禁用'

